(* IEC 61131-3 sources: daoli-st-library/DL_Process (part 39) *)

(* ---- FB_DL_LabelWeekCode.st ---- *)
(*
  Name        : FB_DL_LabelWeekCode
  Category    : DL_Process
  Version     : 1.0.0
  Purpose     : 标签周码/批码打印窗：由年 + 年内日序折算 YYWW 周码，打印请求沿在打印机就绪时发出打印脉冲并锁存周码至请求撤除；/ Label week-code print window: derives a YYWW week code from year and day-of-year, issues a print pulse on request edge when the printer is ready, and latches the code until the request clears
  溯源        : 借 ROADMAP P2（WeekOfYearCalc/DateCoderSync 口径复用），clean-room 实现
  Boundary    : ① 组态闸：年份域 2020..2099 / 年内日序域 1..366 / 打印窗长 > 0 → 锁存故障；
                ② 周码折算：周数 = TRUNC((年内日序 - 1) / 7) + 1（1..53，除子为常量 7，无运行期除零）；
                ③ 打印脉冲 _bPrnC 内部置位 → 段 5 统一出口映射单拍（R187），CASE 内不直写；
                ④ 打印窗计时用 TON 串 ePrint 相位闸（族③），段 0 无 IF 包裹；
                ⑤ nWeekCode 在 eDone 相保持（锁存副本），bPrintReq 撤除沿才回落（族② 保持语义）；
                ⑥ 本件只产生码与脉冲，不驱动打印头（属主边界）。
*)
TYPE E_DL_LwcState :
(
    eIdle  := 0,                             (* 未使能 / Disabled *)
    eReady := 10,                            (* 就绪：等待打印请求（已算码） / Ready *)
    ePrint := 20,                            (* 打印窗进行中 / Printing window *)
    eDone  := 30,                            (* 打印完成（保持周码） / Done, code held *)
    eFault := 90                             (* 故障锁存相 / Fault latched *)
);
END_TYPE

TYPE E_DL_LwcCause :
(
    eNone       := 0,                        (* 无故障成因 / No cause *)
    eCfgIllegal := 1,                        (* 组态非法：年份/日序/窗长越域 / Illegal config *)
    ePhaseBad   := 2                         (* 非法相位兜底 / Illegal phase fallback *)
);
END_TYPE

FUNCTION_BLOCK FB_DL_LabelWeekCode
VAR_INPUT
    nYear     : INT := 2026;                 (* 当前年份，域 2020..2099 [年] / Current year, 2020..2099 *)
    nDayOfYear: INT := 1;                    (* 年内日序（1..366），域 1..366 [日] / Day of year, 1..366 *)
    bPrintReq : BOOL := FALSE;               (* 打印请求电平（上升沿发起）[-] / Print request level *)
    bPrnReady : BOOL := FALSE;               (* 打印机就绪电平 [-] / Printer ready level *)
    tWinLen   : TIME := T#500MS;             (* 打印脉冲窗长，域 > T#0S [ms] / Print pulse window, > 0 *)
    bEnable   : BOOL := TRUE;                (* 使能 [-] / Enable *)
    bReset    : BOOL := FALSE;               (* 复位命令，上升沿清周码与故障 [-] / Reset command *)
END_VAR
VAR_OUTPUT
    nWeekCode : INT;                         (* YYWW 周码（eDone 相保持；低 2 位周数、高位年份后两位）[-] / YYWW week code, held *)
    nWeekNo   : INT;                         (* 年内周数 1..53 [周] / Week number, 1..53 *)
    bPrintPuls: BOOL;                        (* 打印脉冲（窗长电平，tWinLen 定义宽度）[-] / Print pulse level over window *)
    bCodeValid: BOOL;                        (* 周码有效电平（eDone 相为 TRUE）[-] / Code-valid level *)
    eState    : E_DL_LwcState;               (* 状态出口 / State outlet *)
    eCause    : E_DL_LwcCause;               (* 故障成因出口（R190 归因唯一） / Fault cause outlet *)
    bError    : BOOL;                        (* 故障锁存标志 [-] / Fault latch flag *)
END_VAR
VAR
    _eState  : E_DL_LwcState := E_DL_LwcState.eIdle;     (* 内部相位（CASE 唯一写入目标） / Internal phase *)
    _eCause  : E_DL_LwcCause := E_DL_LwcCause.eNone;     (* 故障成因锁存量 / Latched cause *)
    rtReq    : R_TRIG;                       (* 打印请求沿实例，段 0 无条件调用 / Request edge instance *)
    rtReqOff : R_TRIG;                       (* 请求撤除沿实例，段 0 无条件调用 / Request-clear edge instance *)
    rtReset  : R_TRIG;                       (* 复位沿实例，段 0 无条件调用 / Reset edge instance *)
    tonWin   : TON;                          (* 打印脉冲窗计时器（IN 串 ePrint 相位） / Print window timer *)
    _bFault  : BOOL;                         (* 故障锁存位 / Latched fault bit *)
    _bCfgBad : BOOL;                         (* 组态非法当拍量 / Illegal config this scan *)
    _bPrnC   : BOOL;                         (* 打印脉冲窗电平内部量（出口统一映射，R187） / Print-pulse internal level *)
    _nWeekI  : INT;                          (* 周数中间量（折算）[周] / Week number intermediate *)
    _nCodeI  : INT;                          (* 周码中间量（YYWW）[-] / Week code intermediate *)
END_VAR
VAR CONSTANT
    DL_LWC_YMIN  : INT := 2020;              (* 年份域下限 [年] / Year domain floor *)
    DL_LWC_YMAX  : INT := 2099;              (* 年份域上限（YY 码两位十进制安全域）[年] / Year domain ceiling *)
    DL_LWC_DMAX  : INT := 366;               (* 年内日序域上限（含闰年）[日] / Day-of-year domain ceiling *)
    DL_LWC_WMAX  : INT := 53;                (* 周数域上限（折算自洽校验用）[周] / Week number ceiling *)
    DL_LWC_SEVEN : INT := 7;                 (* 周折算除子（常量，无运行期除零）[日/周] / Week divisor *)
    DL_LWC_HUND  : INT := 100;               (* YYWW 折算乘数（常量）[-] / YYWW multiplier *)
END_VAR

(* —— 段 0：当拍判据派生 + 实例无条件刷新（R228A；R_TRIG/TON 全在段 0，无 IF 包裹） —— *)
_bCfgBad := (nYear < DL_LWC_YMIN) OR (nYear > DL_LWC_YMAX)                     (* 年份域闸 / Year gate *)
            OR (nDayOfYear < 1) OR (nDayOfYear > DL_LWC_DMAX)                  (* 日序域闸 / Day-of-year gate *)
            OR NOT (tWinLen > T#0S);                                           (* 窗长正域闸 / Window gate *)
rtReq(CLK := bPrintReq);                                                       (* 请求沿每拍必调 / Request edge every scan *)
rtReqOff(CLK := NOT bPrintReq);                                                (* 请求撤除沿每拍必调 / Request-clear edge every scan *)
rtReset(CLK := bReset);                                                        (* 复位沿每拍必调 / Reset edge every scan *)
tonWin(IN := (_eState = E_DL_LwcState.ePrint) AND bPrintReq, PT := tWinLen);   (* 打印窗计时（串 ePrint 相位闸，族③） / Print timer with phase gate *)

(* —— 段 1：单拍量预清零（R107） —— *)
_bPrnC := FALSE;                                                               (* 打印脉冲内部量预清 / Print-pulse preset *)
bPrintPuls := FALSE;                                                           (* 打印脉冲出口预清 / Print-pulse outlet preset *)
bCodeValid := FALSE;                                                           (* 码有效电平预清 / Code-valid preset *)
_nWeekI := 0;                                                                  (* 周数中间量预清 / Week intermediate preset *)
_nCodeI := 0;                                                                  (* 码中间量预清 / Code intermediate preset *)

(* —— 段 2：复位沿处理（作用域：清故障 + 清周码 + 迁 eIdle，R283 逐项声明） —— *)
IF rtReset.Q THEN
    _bFault := FALSE;                                                          (* 清故障锁存 / Clear fault *)
    _eCause := E_DL_LwcCause.eNone;                                            (* 清成因 / Clear cause *)
    nWeekCode := 0;                                                            (* 清周码出口 / Clear code outlet *)
    nWeekNo := 0;                                                              (* 清周数出口 / Clear week outlet *)
    bCodeValid := FALSE;                                                       (* 清码有效电平 / Clear validity level *)
    _eState := E_DL_LwcState.eIdle;                                            (* 迁未使能相 / Back to idle *)
END_IF

(* —— 段 3：组态故障锁存（锁存至复位沿，R189） —— *)
IF _bCfgBad AND NOT _bFault THEN
    _bFault := TRUE;                                                           (* 锁存故障位 / Latch fault *)
    _eCause := E_DL_LwcCause.eCfgIllegal;                                      (* 成因：组态非法 / Cause: illegal config *)
    _eState := E_DL_LwcState.eFault;                                           (* 同步迁故障相 / Migrate to fault *)
END_IF

(* —— 段 4：CASE 主状态机（ELSE 兜底迁 eFault，红线 6） —— *)
CASE _eState OF
    E_DL_LwcState.eIdle:                                                       (* 未使能：出口确定值 / Disabled *)
        nWeekCode := 0;                                                        (* 失能清周码出口 / Clear code outlet *)
        nWeekNo := 0;                                                          (* 失能清周数出口 / Clear week outlet *)
        bCodeValid := FALSE;                                                   (* 失能清码有效电平 / Clear validity level *)
        IF bEnable AND NOT _bFault THEN
            _eState := E_DL_LwcState.eReady;                                   (* 使能进入就绪 / Enter ready *)
        END_IF
    E_DL_LwcState.eReady:                                                      (* 就绪相：折算周码待打印请求 / Ready *)
        IF NOT bEnable THEN
            _eState := E_DL_LwcState.eIdle;                                    (* 失能回未使能 / Back to idle *)
        ELSE
            _nWeekI := TRUNC(INT_TO_REAL(nDayOfYear - 1) / INT_TO_REAL(DL_LWC_SEVEN)) + 1;   (* 周数折算 = TRUNC((日序-1)/7)+1（除子常量，边界②） / Week number derivation *)
            IF _nWeekI > DL_LWC_WMAX THEN
                _nWeekI := DL_LWC_WMAX;                                        (* 周数上限饱和（最后一次写） / Week ceiling, last write *)
            END_IF
            nWeekNo := _nWeekI;                                                (* 周数出口 / Week outlet *)
            _nCodeI := (nYear MOD DL_LWC_HUND) * DL_LWC_HUND + _nWeekI;        (* YYWW 码 = (年 MOD 100)×100 + 周（乘除均为常量） / YYWW code *)
            nWeekCode := _nCodeI;                                              (* 周码出口（就绪相即为当前码） / Code outlet *)
            IF rtReq.Q AND bPrnReady THEN                                      (* 请求沿 + 就绪：发起打印 / Request edge with ready *)
                _bPrnC := TRUE;                                                (* 打印脉冲内部置位（出口统一映射，R187） / Print-pulse internal *)
                _eState := E_DL_LwcState.ePrint;                               (* 进打印窗相 / To printing *)
            END_IF
        END_IF
    E_DL_LwcState.ePrint:                                                       (* 打印窗相：脉冲电平保持窗长 / Printing *)
        IF NOT bEnable THEN
            _eState := E_DL_LwcState.eIdle;                                    (* 失能回未使能 / Back to idle *)
        ELSE
            _bPrnC := TRUE;                                                    (* 打印窗内脉冲电平保持（窗长由 tonWin 定义） / Pulse level held over window *)
            bCodeValid := TRUE;                                                (* 打印期码有效电平 / Validity level during print *)
            IF rtReqOff.Q THEN                                                 (* 请求撤除沿：提前结束窗 / Request cleared: end window *)
                _eState := E_DL_LwcState.eDone;                                (* 迁完成相（保持周码） / To done *)
            ELSIF tonWin.Q THEN                                                (* 窗长到点：打印完成 / Window elapsed: done *)
                _eState := E_DL_LwcState.eDone;                                (* 迁完成相 / To done *)
            END_IF
        END_IF
    E_DL_LwcState.eDone:                                                       (* 完成相：保持周码至请求撤除后的新请求（族② 保持语义） / Done: hold code *)
        IF NOT bEnable THEN
            _eState := E_DL_LwcState.eIdle;                                    (* 失能回未使能 / Back to idle *)
        ELSIF rtReq.Q THEN                                                     (* 新打印请求沿：重新折算再打印 / New request: re-derive and print *)
            _eState := E_DL_LwcState.eReady;                                   (* 回就绪相重折算 / Back to ready *)
        END_IF
    E_DL_LwcState.eFault:                                                      (* 故障相：冻结保持末值，仅复位沿出 / Fault *)
        ;                                                                      (* 锁存回放（R28） / Replay from latch *)
    ELSE                                                                       (* 非法相位兜底迁安全态 / Illegal phase fallback *)
        _eState := E_DL_LwcState.eFault;                                       (* 迁故障相 / To fault *)
        _bFault := TRUE;                                                       (* 同步锁存 / Latch *)
        _eCause := E_DL_LwcCause.ePhaseBad;                                    (* 成因：非法相位 / Cause: illegal phase *)
END_CASE

(* —— 段 5：出口映射（内部 _b* → 输出，R187；名实双出口，R191） —— *)
bPrintPuls := _bPrnC;                                                          (* 打印脉冲单拍出口 / Print-pulse single-scan outlet *)
bCodeValid := bCodeValid OR (_eState = E_DL_LwcState.eDone);                   (* 码有效电平（打印期与保持期均为 TRUE，族②） / Validity level held in done *)
bError := _bFault;                                                             (* 故障标志镜像 / Fault flag mirror *)
eState := _eState;                                                             (* 状态出口 / State outlet *)
eCause := _eCause;                                                             (* 成因出口 / Cause outlet *)
END_FUNCTION_BLOCK

(* ---- FB_DL_LamEvaGelContent.st ---- *)
(*==============================================================================
 * 组件名称 (Component)  : FB_DL_LamEvaGelContent
 * 所属子库 (Sublibrary) : DL_Process
 * 当前版本 (Version)    : 1.0.0
 * 兼容性 (Platform)     : CODESYS 3.5+ / TwinCAT 3 / 汇川 InoProShop / 施耐德 Machine Expert
 *                         仅依赖 Standard.library（R_TRIG / ABS），零厂商私有库
 * 功能描述 (Function)   : 层压 EVA 交联度估算与合格窗判定。三段工艺换算：
 *                         ① 温度-时间积分 ∫max(0, T - Tref)dt（有效热剂量，
 *                         [°C·min]）；② 线性标定曲线 gel = fGelBase + fKRate·
 *                         Dose（[%]）；③ 合格窗 [fGelLo, fGelHi] 判定。层压
 *                         运行电平控制积分启停。与 Integrator（纯积分）分工：
 *                         本件是积分→标定→判窗三段工艺换算。
 * 来源标签 (Origin)     : ROADMAP §19.2 R12 池（L814），自研 clean-room
 * 边界语义 (Boundary)   : ① 首扫初始化 _bInit（R310：积分类件首拍清剂量）；
 *                         ② 温度 NaN/Inf 拍冻结积分（不累计不判窗）；
 *                         ③ 交联度换算后域钳 [0, 100]（标定外推过冲钳位）；
 *                         ④ 组态闸：基准温度/速率/窗界/扫描秒值域检查 → 故障。
 * 输出语义 (Fallback)   : 【R191】bEnable = FALSE → 积分冻结保持（剂量与交联
 *                         度为资产属性）；eFault 相 → 冻结 + bError = TRUE。
 * 码位     (Codes)      : 按 R297 范式零 16# 码位硬编码；错误出口 BOOL+ENUM(eCause)。
 * 红线自检 (Redline)    : 7 项红线已自检：R1 零全局 ✓｜R2 零物理地址 ✓｜R3 纯 IEC ✓
 *                         R4 除零无涉/NaN 冻结/钳位/组态闸 ✓｜R5 双语同行注释 ✓
 *                         R6 CASE 带 ELSE 兜底迁 eFault ✓｜R7 R_TRIG 段 0 无条件刷新 ✓
 * 验收向量 (Acceptance) : V1 T=150 恒定、Tref=140、fScanS=1.0、fKRate=0.02：
 *                         600 s 后 Dose = 600·10/60 = 100 [°C·min]，
 *                         gel = 基准 20 + 0.02·100 = 22.0 [%]；
 *                         V2 T <= Tref 全程 → Dose=0，gel=基准（不超下界）；
 *                         V3 gel > 100 外推过冲 → 钳 100（边界③）。
 * 修订历史 (Revision)   : 2026-11-20  v1.0.0  R51 首版（批 2 · 序号 10）
 *==============================================================================*)
TYPE E_DL_LgcState :
(
    eIdle  := 0,                             (* 待使能 / Idle *)
    eCalc  := 10,                            (* 积分与判窗运行 / Calc run *)
    eFault := 90                             (* 故障锁存相 / Fault latched phase *)
);
END_TYPE

TYPE E_DL_LgcCause :
(
    eNone       := 0,                        (* 无故障成因 / No cause *)
    eCfgIllegal := 1,                        (* 组态非法：基准/速率/窗界越域 / Illegal config *)
    ePhaseBad   := 2                         (* 非法相位兜底 / Illegal phase fallback *)
);
END_TYPE

FUNCTION_BLOCK FB_DL_LamEvaGelContent
VAR_INPUT
    fTempC    : LREAL := 25.0;               (* 层压温度 [°C] / Lamination temperature *)
    fTempRef  : LREAL := 140.0;              (* 交联基准温度（低于不累计），域 > 0 [°C] / Reference temperature *)
    fKRate    : LREAL := 0.02;               (* 标定斜率，域 > 0 [%/(°C·min)] / Calibration rate *)
    fGelBase  : LREAL := 20.0;               (* 交联度基准截距，域 [0,100] [%] / Base gel content *)
    fGelLo    : LREAL := 75.0;               (* 合格窗下限，域 < fGelHi [%] / Gel window lower *)
    fGelHi    : LREAL := 95.0;               (* 合格窗上限，域 > fGelLo [%] / Gel window upper *)
    fScanS    : LREAL := 1.0;                (* 扫描周期秒值，域 > 1E-6 [s] / Scan period seconds *)
    bProcRun  : BOOL := FALSE;               (* 层压运行电平（积分启停）[-] / Process run level *)
    bEnable   : BOOL := TRUE;                (* 使能 [-] / Enable *)
    bReset    : BOOL := FALSE;               (* 复位命令，上升沿清剂量与输出 [-] / Reset command *)
END_VAR
VAR_OUTPUT
    fDose     : LREAL;                       (* 有效热剂量 [°C·min] / Effective thermal dose *)
    fGelPct   : LREAL;                       (* 交联度估算（钳 0..100）[%] / Gel content estimate *)
    bGelOk    : BOOL;                        (* 合格窗判定（窗口内）[-] / Gel-in-window verdict *)
    eState    : E_DL_LgcState;               (* 状态出口 / State outlet *)
    eCause    : E_DL_LgcCause;               (* 故障成因出口 / Fault cause outlet *)
    bError    : BOOL;                        (* 故障锁存标志 [-] / Fault latch flag *)
END_VAR
VAR
    _eState  : E_DL_LgcState := E_DL_LgcState.eIdle;      (* 内部相位（CASE 唯一写入目标） / Internal phase *)
    _eCause  : E_DL_LgcCause := E_DL_LgcCause.eNone;      (* 故障成因锁存量 / Latched cause *)
    rtReset  : R_TRIG;                       (* 复位沿实例，段 0 无条件调用 / Reset edge instance *)
    _fDose   : LREAL;                        (* 剂量积分锁存 [°C·min] / Dose integrator latch *)
    _fGel    : LREAL;                        (* 交联度派生量 [%] / Gel derived *)
    _bTempBad: BOOL;                         (* 温度非有限当拍量 [-] / Non-finite temperature *)
    _bInit   : BOOL := FALSE;                (* 首扫初始化标志（R310）[-] / First-scan init flag *)
    _bFault  : BOOL;                         (* 故障锁存位 / Latched fault bit *)
    _bCfgBad : BOOL;                         (* 组态非法当拍量 / Illegal config this scan *)
END_VAR
VAR CONSTANT
    DL_LGC_EPS : LREAL := 1.0E-6;            (* 秒值判零容差 [s] / Seconds epsilon *)
    DL_LGC_MIN : LREAL := 60.0;              (* 秒 → 分换算常量 [s/min] / Seconds per minute *)
    DL_LGC_GMAX: LREAL := 100.0;             (* 交联度物理上限 [%] / Gel physical max *)
    DL_LGC_INF : LREAL := 1.0E30;            (* Inf 差判兜底量纲界 [—] / Inf diff guard *)
END_VAR

(* —— 段 0：当拍判据派生 + 实例无条件刷新（R228A） —— *)
_bCfgBad := (fTempRef <= 0.0) OR (fKRate <= 0.0) OR (fGelBase < 0.0) OR (fGelBase > DL_LGC_GMAX)
            OR (fGelLo >= fGelHi) OR (fScanS <= DL_LGC_EPS);   (* 组态闸（R151 全引脚 + 窗界序） / Config gate *)
rtReset(CLK := bReset);                      (* 复位沿每拍必调 / Reset edge every scan *)
_bTempBad := (fTempC <> fTempC) OR ((fTempC - fTempC) <> (fTempC - fTempC))
            OR (ABS(fTempC) > DL_LGC_INF);   (* 温度 NaN 自反 + Inf 差判 + 量纲兜底 / Non-finite temperature *)

(* —— 段 1：首扫初始化（R310：积分类件首拍清剂量，与复位沿同款） —— *)
IF NOT _bInit THEN
    _fDose := 0.0;                           (* 首拍剂量清零 / First-scan dose clear *)
    _fGel := fGelBase;                       (* 首拍交联度取基准 / First-scan gel base *)
    _bInit := TRUE;                          (* 置初始化完成 / Set init done *)
END_IF
_fGel := 0.0;                                (* 交联度当拍量预清（每拍全路径派生，R285） / Gel preset *)
bGelOk := FALSE;                             (* 判窗预清（全路径赋值） / Verdict preset *)

(* —— 段 2：复位沿处理（作用域：清故障 + 清剂量积分 + 清输出 + 迁 eIdle，R283 逐项声明） —— *)
IF rtReset.Q THEN
    _bFault := FALSE;                        (* 清故障锁存 / Clear fault *)
    _eCause := E_DL_LgcCause.eNone;          (* 清成因 / Clear cause *)
    _fDose := 0.0;                           (* 清剂量积分 / Clear dose *)
    fDose := 0.0;                            (* 清剂量出口 / Clear dose outlet *)
    fGelPct := fGelBase;                     (* 交联度回基准 / Gel back to base *)
    _eState := E_DL_LgcState.eIdle;          (* 迁待机相 / Back to idle *)
END_IF

(* —— 段 3：组态闸故障锁存（R45 配对；锁存至复位沿，R189） —— *)
IF _bCfgBad AND NOT _bFault THEN
    _bFault := TRUE;                         (* 锁存故障位 / Latch fault *)
    _eCause := E_DL_LgcCause.eCfgIllegal;    (* 成因：组态非法 / Cause: illegal config *)
    _eState := E_DL_LgcState.eFault;         (* 同步迁故障相 / Migrate to fault *)
END_IF

(* —— 段 4：CASE 主状态机（ELSE 兜底迁 eFault，红线 6） —— *)
CASE _eState OF
    E_DL_LgcState.eIdle:                     (* 待机相 / Idle *)
        IF bEnable AND NOT _bFault AND NOT _bTempBad THEN
            _eState := E_DL_LgcState.eCalc;  (* 进入计算 / Enter calc *)
        END_IF
    E_DL_LgcState.eCalc:                     (* 计算相：积分 + 标定 + 判窗 / Calc *)
        IF NOT bEnable THEN
            _eState := E_DL_LgcState.eIdle;  (* 失能回待机（剂量冻结保持，R191 声明） / Back to idle, dose held *)
        ELSIF bProcRun AND (NOT _bTempBad) THEN   (* 运行电平 + 温度有限才积分 / Integrate when running *)
            IF fTempC > fTempRef THEN        (* 有效热剂量：仅高于基准累计 / Dose above reference *)
                _fDose := _fDose + (fTempC - fTempRef) * fScanS / DL_LGC_MIN;   (* 增量 = ΔT·dt/60 [°C·min]，除子常量 60 无除零 / Dose increment *)
            END_IF
        END_IF                               (* 温度坏值/停运拍：积分冻结（边界②） / Freeze on bad temp *)
        _fGel := fGelBase + fKRate * _fDose; (* 标定曲线换算（乘法无除零） / Calibration transform *)
        IF _fGel < 0.0 THEN
            _fGel := 0.0;                    (* 下界钳位 / Lower clamp *)
        ELSIF _fGel > DL_LGC_GMAX THEN
            _fGel := DL_LGC_GMAX;            (* 上界钳位（外推过冲兜底，边界③） / Upper clamp *)
        END_IF
        IF (_eState = E_DL_LgcState.eCalc) AND (NOT _bTempBad) THEN   (* 判窗仅运行域有效拍 / Verdict in valid scans *)
            fDose := _fDose;                 (* 剂量出口刷新 / Dose outlet *)
            fGelPct := _fGel;                (* 交联度出口刷新 / Gel outlet *)
            IF _fGel < fGelLo THEN
                bGelOk := FALSE;             (* 低于窗 / Below window *)
            ELSIF _fGel > fGelHi THEN
                bGelOk := FALSE;             (* 高于窗 / Above window *)
            ELSE
                bGelOk := TRUE;              (* 窗内（IF 链带 ELSE 兜底，R285） / In window *)
            END_IF
        END_IF
    E_DL_LgcState.eFault:                    (* 故障相：冻结保持，仅复位沿出 / Fault *)
        ;                                    (* 锁存回放（R28） / Replay from latch *)
    ELSE                                     (* 非法相位兜底迁安全态 / Illegal phase fallback *)
        _eState := E_DL_LgcState.eFault;     (* 迁故障相 / To fault *)
        _bFault := TRUE;                     (* 同步锁存 / Latch *)
        _eCause := E_DL_LgcCause.ePhaseBad;  (* 成因：非法相位 / Cause: illegal phase *)
END_CASE

(* —— 段 5：出口映射（bError/eState 同源，R191） —— *)
bError := _bFault;                           (* 故障标志镜像 / Fault flag mirror *)
eState := _eState;                           (* 状态出口 / State outlet *)
eCause := _eCause;                           (* 成因出口 / Cause outlet *)
END_FUNCTION_BLOCK

(* ---- FB_DL_LamHeaterZoneSync.st ---- *)
//==============================================================================
// 功能块：FB_DL_LamHeaterZoneSync ｜ 中文名称：层压机加热板多温区同步跟随
// 所属子库：DL_Process ｜ 版本：v1.0.0 ｜ 兼容：CODESYS V3.5+ / TwinCAT 3 / 汇川 InoProShop
// 功能描述：层压机加热板多温区同步监视——计算有效温区两两最大区差与
//           最差温差对，区差超阈值经确认窗（防瞬态抖动）判失步故障；
//           链速参与跟随语义（链速为 0 时跟随斜率冻结，不除零）。
// 开源溯源 (Origin)：道莅原创实现（参考光伏组件层压机工程惯例 分类与参数域）
// 单位表：T[°C] / 区差[K] / 链速[mm/s] / 确认窗[ms] / 温区下标[区]
// 错误码表：16#0005_01E6 信息级（非有限温区剔除声明，不置 bError）/
//           16#0005_01E7 信息级（区数上限已钳位 8，不置 bError）/
//           16#0005_031E 故障级（区差超限经确认窗确认，置 bError）/
//           16#0005_031F 故障级（有效区数 < 2 无法判区差，置 bError）/
//           16#0005_0320 故障级兜底（置 bError）
// 状态机：N/A（阈值确认窗 + 电平逻辑，无相位状态机；故障经确认窗后以
//           bSyncOk 电平与 031E 表达，原因消失自动恢复，无锁存）
// 边界行为：① 区差 > 阈值持续确认窗 → 故障 031E + bSyncOk := FALSE
//           （R13 AhuDamperStuckDiag 确认窗范式复用）；② 任一温区非有限
//           → 该区剔除出区差统计 + 信息 01E6；有效区数 < 2 → 故障 031F；
//           ③ 链速为 0 → 跟随斜率冻结（不除零），区差统计不受影响；
//           ④ 区数上限钳 8 + 信息 01E7（接口字面量上界 8 与 DL_ZONE_MAX
//           同源，一致性由本件承担验证责任）；⑤ 非使能时输出冻结为零
//           值并 bValid := FALSE（不静默沿用旧差值）。
// 依赖纪律：仅 Standard.library；零跨层调用（两两区差为 O(n²) 遍历的
//           监视语义，非统计算法复制，头注释声明此设计取舍）。
// 修订历史：v1.0.0 2026-11-17 首版（R23 派单 · ROADMAP 光伏 P1 §416）
//==============================================================================

FUNCTION_BLOCK FB_DL_LamHeaterZoneSync
VAR_INPUT
    aZoneTempC    : ARRAY[1..8] OF LREAL;   // 各温区实测 [摄氏度]，下标 1..8，超编路填 0 且不计 / Measured zone temperatures [degC], index 1..8
    uZoneCount    : UINT;                   // 实际温区数 [区]，有效域 0..8，> 8 钳位 / Actual zone count [zones], 0..8, clamped above
    fZoneDiffMaxK : LREAL := 5.0;           // 区差阈值 [K]，须 > 0 / Zone-difference threshold [K], must be > 0
    fBeltSpeedMmS : LREAL;                  // 链速 [毫米/秒]，0 = 停链（跟随冻结） / Belt speed [mm/s], zero = stopped, follow frozen
    bEnable       : BOOL;                   // 使能 [—] / Enable
    bReset        : BOOL;                   // 故障复位 [—]，清除确认窗 / Fault reset, clears the confirm window
END_VAR
VAR_OUTPUT
    fMaxZoneDiffK : LREAL;                  // 当拍最大区差 [K] / Maximum zone difference this scan [K]
    bSyncOk       : BOOL;                   // 同步正常 [—] / Synchronization OK
    uWorstPairA   : UINT;                   // 最大温差对 A 区下标 [区] / Worst pair index A [zone]
    uWorstPairB   : UINT;                   // 最大温差对 B 区下标 [区] / Worst pair index B [zone]
    eErr          : UDINT;                  // 错误码，0 = 无错 / Error code, 0 = no error
    bError        : BOOL;                   // 故障级标志，仅故障级错误置位 / Fault-class flag, set only on fault-level codes
    bValid        : BOOL;                   // 输出可用标志 / Outputs usable flag
END_VAR
VAR
    fbConfirm     : TON;                    // 区差超限确认窗，段 6 无条件刷新 [ms] / Zone-diff confirm window
    _uCountEff    : UINT;                   // 钳位后的生效区数 [区] / Effective clamped zone count
    _uValidZones  : UINT;                   // 非有限剔除后的有效区数 [区] / Valid zone count after culling
    _uI           : UINT;                   // 外层遍历下标 [区] / Outer loop index
    _uJ           : UINT;                   // 内层遍历下标 [区] / Inner loop index
    _fDiff        : LREAL;                  // 当前对区差 [K] / Current pair difference [K]
    _bInit        : BOOL := FALSE;          // 首扫标志，初值 FALSE 取非判定 / First-scan flag, tested negated
    _bCullInfo    : BOOL;                   // 非有限剔除信息当拍标志 / Cull info flag of this scan
    _bClampInfo   : BOOL;                   // 区数钳位信息当拍标志 / Clamp info flag of this scan
    _bIllegal     : BOOL;                   // 非法输入标志（阈值非有限/<= 0） / Illegal input flag
END_VAR
VAR CONSTANT
    DL_ZONE_MAX   : UINT  := 8;             // 温区上限 [区]，与接口字面量上界 8 同源，改动须同步 / Zone ceiling [zones], same source as the literal bound 8, change both together
    DL_LAM_INF    : LREAL := 1.7976931348623157E308; // LREAL 幅值上限 / LREAL magnitude ceiling
    DL_LAM_CONFIRM: TIME  := T#10S;         // 区差超限确认窗 [ms]（R13 范式） / Zone-diff confirm window [ms], R13 pattern
END_VAR

(*------------------------------------------------------------------------------
 * 段 1｜每拍预置：输出先算后出，单拍标志预清零
 *      Outputs computed per scan, one-shot flags pre-cleared
 *-----------------------------------------------------------------------------*)
fMaxZoneDiffK := 0.0;                       // 最大区差预置零 / Max difference preset zero
bSyncOk       := FALSE;                     // 同步正常预置 FALSE / Sync OK preset FALSE
uWorstPairA   := 0;                         // 最差对 A 预置零 / Worst A preset zero
uWorstPairB   := 0;                         // 最差对 B 预置零 / Worst B preset zero
eErr          := 16#0000_0000;              // 错误码每拍重算 / Error code recomputed
bError        := FALSE;                     // 故障标志每拍重算 / Fault flag recomputed
bValid        := FALSE;                     // 可用标志每拍重算 / Usable flag recomputed
_bCullInfo    := FALSE;                     // 剔除信息预清零 / Cull info pre-cleared
_bClampInfo   := FALSE;                     // 钳位信息预清零 / Clamp info pre-cleared
_bIllegal     := FALSE;                     // 非法输入预清零 / Illegal input pre-cleared

(*------------------------------------------------------------------------------
 * 段 2｜首扫初始化
 *      First-scan initialisation
 *-----------------------------------------------------------------------------*)
IF NOT _bInit THEN
    _uCountEff := 0;                        // 生效区数从零起步 / Effective count starts at zero
    _bInit     := TRUE;                     // 首扫只做一次 / The first scan runs once
END_IF

(*------------------------------------------------------------------------------
 * 段 3｜组态与输入防御闸（阈值非法 / 区数钳位）
 *      Configuration and input defense gates
 *-----------------------------------------------------------------------------*)
IF (fZoneDiffMaxK <> fZoneDiffMaxK) OR (ABS(fZoneDiffMaxK) > DL_LAM_INF) OR (fZoneDiffMaxK <= 0.0) THEN
    _bIllegal := TRUE;                      // 阈值非法（031F 无法判差的同类防御，R90 精神） / Illegal threshold
END_IF
IF (fBeltSpeedMmS <> fBeltSpeedMmS) OR (ABS(fBeltSpeedMmS) > DL_LAM_INF) THEN
    _bIllegal := TRUE;                      // 链速非有限防御 / Non-finite belt speed
END_IF
IF uZoneCount > DL_ZONE_MAX THEN
    _uCountEff := DL_ZONE_MAX;              // 区数钳位到 8 / Zone count clamped to 8
    _bClampInfo := TRUE;                    // 钳位信息置位 / Clamp info raised
ELSE
    _uCountEff := uZoneCount;               // 合法区数原值生效 / Valid count applied as-is
END_IF

(*------------------------------------------------------------------------------
 * 段 4｜两两区差扫描（非有限区剔除 + 最差对记录）
 *      Pairwise scan with non-finite culling and worst-pair recording
 *-----------------------------------------------------------------------------*)
_uValidZones := 0;                          // 有效区数清零 / Valid count cleared
FOR _uI := 1 TO _uCountEff DO
    IF _uI <= DL_ZONE_MAX THEN              // 二次闸：越界结构性不可能 / Secondary gate, out-of-bounds impossible
        IF (aZoneTempC[_uI] <> aZoneTempC[_uI]) OR (ABS(aZoneTempC[_uI]) > DL_LAM_INF) THEN
            _bCullInfo := TRUE;             // 非有限区剔除声明 / Non-finite zone culled
        ELSE
            _uValidZones := _uValidZones + 1; // 有效区计数递增 / Valid count increment
        END_IF
        FOR _uJ := _uI + 1 TO _uCountEff DO
            IF _uJ <= DL_ZONE_MAX THEN      // 二次闸 / Secondary gate
                IF (aZoneTempC[_uI] <> aZoneTempC[_uI]) OR (ABS(aZoneTempC[_uI]) > DL_LAM_INF)
                   OR (aZoneTempC[_uJ] <> aZoneTempC[_uJ]) OR (ABS(aZoneTempC[_uJ]) > DL_LAM_INF) THEN
                    (* 任一侧非有限：本对剔除，不计入区差 / Either side non-finite, the pair is culled *)
                    _fDiff := 0.0;          // 本对区差按零计（不参与最差对竞争） / Pair difference counted as zero
                ELSE
                    _fDiff := ABS(aZoneTempC[_uI] - aZoneTempC[_uJ]); // 当前对区差 [K] / Current pair difference [K]
                    IF _fDiff > fMaxZoneDiffK THEN
                        fMaxZoneDiffK := _fDiff; // 更新最大区差 / Update the max difference
                        uWorstPairA := _uI;  // 记录最差对 A / Record worst pair A
                        uWorstPairB := _uJ;  // 记录最差对 B / Record worst pair B
                    END_IF
                END_IF
            END_IF
        END_FOR
    END_IF
END_FOR

(*------------------------------------------------------------------------------
 * 段 5｜确认窗无条件刷新（R40：CASE 之外每拍必调）
 *      Confirm window refreshed unconditionally per R40
 *-----------------------------------------------------------------------------*)
fbConfirm(IN := bEnable AND (NOT _bIllegal) AND (_uValidZones >= 2)
              AND (NOT bReset) AND (fMaxZoneDiffK > fZoneDiffMaxK), PT := DL_LAM_CONFIRM); // 区差超限确认窗（bReset 电平拦截断窗复位） / Zone-diff confirm window, bReset breaks the input to reset

(*------------------------------------------------------------------------------
 * 段 6｜出口与码位（链速为 0 时跟随斜率冻结——本件无斜率输出引脚，
 *       跟随联动由调用方按 fBeltSpeedMmS = 0 自行冻结，边界声明）
 *      Outlet and codes, belt-speed freeze declared for the caller
 *-----------------------------------------------------------------------------*)
IF (NOT bEnable) OR _bIllegal THEN
    bValid := FALSE;                        // 未使能或输入非法：输出不可用 / Not enabled or illegal input, outputs unusable
ELSIF _uValidZones < 2 THEN
    eErr   := 16#0005_031F;                 // 故障级：有效区数 < 2 无法判区差 / Fault: fewer than two valid zones
    bError := TRUE;                         // 置故障标志（R45 配对） / Raise the fault flag
    bValid := FALSE;                        // 输出不可用 / Outputs unusable
ELSIF fbConfirm.Q THEN
    eErr   := 16#0005_031E;                 // 故障级：区差超限经确认窗确认 / Fault: zone difference confirmed
    bError := TRUE;                         // 置故障标志 / Raise the fault flag
    bSyncOk := FALSE;                       // 失步声明 / Desynchronization declared
    bValid := TRUE;                         // 判定结果本身可用 / The verdict itself is usable
ELSE
    bSyncOk := TRUE;                        // 同步正常 / Synchronized
    IF _bCullInfo THEN
        eErr := 16#0005_01E6;               // 信息级：非有限温区已剔除 / Info: non-finite zones culled
    END_IF
    IF _bClampInfo THEN
        eErr := 16#0005_01E7;               // 信息级：区数已钳位 8 / Info: zone count clamped to 8
    END_IF
    bValid := TRUE;                         // 输出可用 / Outputs usable
END_IF
END_FUNCTION_BLOCK

(* ---- FB_DL_LaminatorTempProfile.st ---- *)
(*
  FB_DL_LaminatorTempProfile  —  层压机多温区配方曲线跟随 / Laminator multi-zone temperature profile
  分类 Category : DL_Process
  码位 Code     : 16#06_0_8D
  版本 Version  : 1.0.0
  溯源 Source   : LGF Technology 语义借鉴 · clean-room 实现，仅借分类/参数域/命名，未复制源码
  功能 Function : 1) 每温区按「升温 → 保温 → 降温」三段配方跟随（复用 FB_DL_RampSoakProfile 多实例按温区展开）；
                  2) 全部温区过各自终点窗才置 bProfileDone（单区完成不算完成）；
                  3) 任一温区实测温度无效：该区冻结判定保持末次设定，其余区继续。
  边界 Boundary : ① 段表非法（斜率 <= 0 折算斜坡时间 <= 0、保温时长 < 0、温区数越界）出厂报码；
                  ② 实测温度非有限判 NE43 无效：该温区冻结判定并置信息码，禁塞伪值；
                  ③ 段切换沿冻结一拍防设定阶跃（切换拍不更新区设定输出）；
                  ④ 超时未达窗升级为段故障（锁存），不死等；
                  ⑤ 输出三行同向：区段号 → 区设定 → 完成标志。
  依赖 Depends  : FB_DL_RampSoakProfile × DL_LAM_ZMAX（设定源实例，每拍无条件调用）
  职责边界 Note : 与 FB_DL_CvdTempRamp 同用 RampSoakProfile，但本件面向层压机三段真空/加压
                  配方（段数固定 3、有 bHoldActive 保温保持出口），CVD 件面向多段 Ramp/Soak +
                  均匀性判据，二者行业参数集与判据分立，互不替代。

  码表 Error codes（本件子码步进 16#10，避让邻件码位）:
    16#0002_068D 故障级：段表组态非法（温区数越界 / 斜坡或保温时长 < 0 / 目标温度非有限）
    16#0002_069D 故障级：段超时（保温段计时超限时仍未达窗，锁存需复位）
    16#0002_06AD 信息级：某温区实测温度无效，该区判定已冻结（不置 bError）
*)

TYPE E_DL_LtpPhase :
(
    eIdle    := 0,   // 空闲 / Idle
    eRun     := 10,  // 曲线跟随中 / Profile running
    eDone    := 20,  // 全区完成 / All zones done
    eFrozen  := 30,  // 全部温区无效冻结 / All zones frozen by invalid feedback
    eFault   := 90   // 段故障锁定 / Segment fault locked
);
END_TYPE

FUNCTION_BLOCK FB_DL_LaminatorTempProfile
VAR_INPUT
    bStart        : BOOL;                           // 启动指令，上升沿生效 / Profile start, edge
    bHold         : BOOL;                           // 外部保持（暂停整条曲线）/ External hold
    bReset        : BOOL;                           // 复位，上升沿清段故障 / Reset, clears segment fault
    nZoneCount    : INT := 3;                       // 温区数 [区]，1..DL_LAM_ZMAX / Zone count
    aTgtRampC     : ARRAY[1..4] OF REAL;            // 升温段目标 [°C] × 区 / Ramp segment target [degC] per zone
    aTgtSoakC     : ARRAY[1..4] OF REAL;            // 保温段目标 [°C] × 区 / Soak segment target [degC] per zone
    aTgtCoolC     : ARRAY[1..4] OF REAL;            // 降温段目标 [°C] × 区 / Cool segment target [degC] per zone
    aTempActC     : ARRAY[1..4] OF REAL;            // 各温区实测温度 [°C] / Measured zone temperature [degC]
    tRampUp       : TIME := T#600S;                 // 升温段斜坡时间 [s] / Ramp-up duration
    tSoak         : TIME := T#900S;                 // 保温段保持时间 [s] / Soak duration
    tCoolDown     : TIME := T#600S;                 // 降温段斜坡时间 [s] / Cool-down duration
    fEndWinK      : REAL := 3.0;                    // 终点窗半宽 [K]，域 > 0 / End window half width [K]
    fEps          : REAL := 1.0E-6;                 // 浮点判零容差 [1] / Floating zero tolerance
END_VAR
VAR_OUTPUT
    afZoneSpC     : ARRAY[1..4] OF REAL;            // 各温区设定输出 [°C] / Zone setpoint output [degC]
    anZoneSeg     : ARRAY[1..4] OF INT;             // 各温区当前段号 1..3 / Active segment per zone
    bProfileDone  : BOOL;                           // 全部温区过终点窗 / All zones past end window
    bHoldActive   : BOOL;                           // 保温段激活标志（任一区在保温段）/ Any zone in soak segment
    bError        : BOOL;                           // 故障标志，与故障级码配对 / Fault flag paired with fault codes
    uErrorId      : UDINT;                          // 事件码，0 = 无事件 / Event code, 0 = none
    eStateOut     : E_DL_LtpPhase;                  // 状态机当前态，段尾单点映射 / Phase mapped at tail
END_VAR
VAR
    _eState       : E_DL_LtpPhase := E_DL_LtpPhase.eIdle;  // 内部状态 / Internal state
    afbRs         : ARRAY[1..4] OF FB_DL_RampSoakProfile;  // 每温区一条曲线实例（无条件调用）/ Per-zone profile instance
    rtrStart      : R_TRIG;                         // 启动沿 / Start edge
    rtrReset      : R_TRIG;                         // 复位沿 / Reset edge
    abZoneFrozen  : ARRAY[1..4] OF BOOL;            // 温区冻结掩码（实测无效）/ Zone frozen mask
    abZoneDone    : ARRAY[1..4] OF BOOL;            // 温区过终点窗掩码 / Zone end-window mask
    abSegChgPrev  : ARRAY[1..4] OF BOOL;            // 上拍段切换沿（冻结一拍用）/ Previous segment-change edge
    bCfgOk        : BOOL;                           // 组态合法标志 / Configuration valid
    bZoneOk       : BOOL;                           // 本拍温度数组有效（逐区判定）/ Zone validity this scan
    bAnyFrozen    : BOOL;                           // 存在冻结区 / Any zone frozen
    bAllInvalid   : BOOL;                           // 全部温区无效 / All zones invalid
    nZ            : INT;                            // 温区遍历索引 / Zone loop index
    nSegMax       : INT;                            // 全区最大段号（输出口径）/ Max segment across zones
    uFault        : UDINT;                          // 锁存故障码 / Latched fault code
    uInfo         : UDINT;                          // 信息级码 / Information code
    bTonArmed     : BOOL;                           // 段超时定时器装载条件 / Segment timeout arming condition
END_VAR
VAR CONSTANT
    DL_LAM_ZMAX   : INT := 4;                       // 温区数上限 [区] / Zone count upper bound
    DL_LAM_INFMAX : REAL := 1.0E30;                 // 温度有限值幅值上限 [°C] / Temperature finite bound [degC]
END_VAR

(* === 段 0 · 实例刷新 === *)
rtrStart(CLK := bStart);                          // 每拍刷新启动沿
rtrReset(CLK := bReset);                          // 每拍刷新复位沿

(* === 段 1 · 组态闸 === *)
bCfgOk := (nZoneCount >= 1) AND (nZoneCount <= DL_LAM_ZMAX)    // 温区数域闸
          AND (TIME_TO_REAL(tRampUp) > 0.0)                     // 升温时长 > 0（斜率合法性由时长承载）
          AND (TIME_TO_REAL(tCoolDown) > 0.0) AND (TIME_TO_REAL(tSoak) >= 0.0)
          AND (fEndWinK > fEps);                                // 终点窗半宽正域
FOR nZ := 1 TO DL_LAM_ZMAX DO
    bCfgOk := bCfgOk AND (aTgtRampC[nZ] = aTgtRampC[nZ])        // 目标温度 NaN 自反
              AND (aTgtSoakC[nZ] = aTgtSoakC[nZ]) AND (aTgtCoolC[nZ] = aTgtCoolC[nZ])
              AND (ABS(aTgtRampC[nZ]) < DL_LAM_INFMAX)          // 幅值域闸（仅组态域，实测另行判定）
              AND (ABS(aTgtSoakC[nZ]) < DL_LAM_INFMAX) AND (ABS(aTgtCoolC[nZ]) < DL_LAM_INFMAX);
END_FOR
IF NOT bCfgOk THEN
    uFault := 16#0002_068D;                       // 故障级：段表组态非法
END_IF
IF rtrReset.Q AND bCfgOk THEN
    uFault := 16#0000;                            // 复位沿清段故障锁存（解除路径可达）
    FOR nZ := 1 TO DL_LAM_ZMAX DO
        abZoneDone[nZ] := FALSE;                  // 完成掩码同步复位
        abZoneFrozen[nZ] := FALSE;                // 冻结掩码同步复位
    END_FOR
END_IF
uInfo := 16#0000;                                 // 信息码每拍清零

(* === 段 2 · 逐温区实例调用（无条件）与实测域闸 === *)
bAnyFrozen := FALSE;                              // 冻结汇总先清
bAllInvalid := TRUE;                              // 全无效假设先置
FOR nZ := 1 TO DL_LAM_ZMAX DO
    bZoneOk := (aTempActC[nZ] = aTempActC[nZ]) AND (ABS(aTempActC[nZ]) < DL_LAM_INFMAX);  // NaN 自反 + 幅值闸
    IF bZoneOk THEN
        abZoneFrozen[nZ] := FALSE;                // 该区恢复有效
        abZoneDone[nZ] := abZoneDone[nZ] OR (ABS(aTempActC[nZ] - aTgtCoolC[nZ]) <= fEndWinK + fEps);  // 过终点窗判定（保持型）
        afbRs[nZ](bStart := rtrStart.Q,           // 启动沿下发
                  bHold := bHold OR abZoneFrozen[nZ],   // 外部保持或该区无效冻结（实例内冻结计时）
                  fTrackValue := aTempActC[nZ],   // 无效恢复后无扰回投基准
                  bTrack := FALSE,                // 有效区不跟踪（跟踪入口仅供无效恢复衔接）
                  nSegCount := 3,                 // 固定三段：升温/保温/降温
                  aTarget[1] := aTgtRampC[nZ],    // 段 1 目标：升温
                  aTarget[2] := aTgtSoakC[nZ],    // 段 2 目标：保温
                  aTarget[3] := aTgtCoolC[nZ],    // 段 3 目标：降温
                  aRampTime[1] := tRampUp,        // 段 1 斜坡时间
                  aRampTime[2] := T#0S,           // 段 2 阶跃直达保温目标（保温由时长承载）
                  aRampTime[3] := tCoolDown,      // 段 3 斜坡时间
                  aSoakTime[1] := T#0S,           // 升温到位即切段
                  aSoakTime[2] := tSoak,          // 保温时长
                  aSoakTime[3] := T#0S,           // 降温到位即完成
                  bLoopProfile := FALSE,          // 单次配方不循环
                  bReset := rtrReset.Q);          // 复位沿透传
        IF afbRs[nZ].bSegChange THEN
            abSegChgPrev[nZ] := TRUE;             // 段切换沿：下一拍冻结一拍防设定阶跃
        ELSE
            abSegChgPrev[nZ] := FALSE;            // 非切换拍清标记
        END_IF
        IF NOT abSegChgPrev[nZ] THEN
            afZoneSpC[nZ] := afbRs[nZ].fSetpoint; // 非冻结拍：区设定跟随曲线
        END_IF                                    // 冻结拍：保持上拍设定（防阶跃）
        anZoneSeg[nZ] := afbRs[nZ].nSegAct;       // 段号输出
    ELSE
        abZoneFrozen[nZ] := TRUE;                 // 该区判定冻结（不塞伪值）
        uInfo := 16#0002_06AD;                    // 信息级：温区实测无效该区冻结
        afbRs[nZ](bStart := FALSE, bHold := TRUE, bReset := FALSE,   // 实例仍无条件调用：保持态
                  fTrackValue := aTempActC[nZ], bTrack := TRUE,      // 跟踪入口挂无效值会被实例自身域闸拒绝
                  nSegCount := 3, aTarget[1] := aTgtRampC[nZ], aTarget[2] := aTgtSoakC[nZ],
                  aTarget[3] := aTgtCoolC[nZ], aRampTime[1] := tRampUp, aRampTime[2] := T#0S,
                  aRampTime[3] := tCoolDown, aSoakTime[1] := T#0S, aSoakTime[2] := tSoak,
                  aSoakTime[3] := T#0S, bLoopProfile := FALSE);
        anZoneSeg[nZ] := afbRs[nZ].nSegAct;       // 段号照透传（判定冻结但显示不冻结）
    END_IF
    bAnyFrozen := bAnyFrozen OR abZoneFrozen[nZ]; // 汇总冻结
    bAllInvalid := bAllInvalid AND (NOT bZoneOk); // 汇总全无效
END_FOR

(* === 段 3 · 主状态机（ENUM + CASE，含 ELSE 兜底）=== *)
CASE _eState OF
E_DL_LtpPhase.eIdle :
    bProfileDone := FALSE;                        // 空闲未完成
    bHoldActive := FALSE;                         // 空闲无保温
    IF uFault <> 16#0000 THEN
        _eState := E_DL_LtpPhase.eFault;          // 故障优先
    ELSIF bAllInvalid AND bCfgOk THEN
        _eState := E_DL_LtpPhase.eFrozen;         // 全区无效进冻结
    ELSIF (afbRs[1].nSegAct > 0) OR (afbRs[2].nSegAct > 0)
      OR (afbRs[3].nSegAct > 0) OR (afbRs[4].nSegAct > 0) THEN
        _eState := E_DL_LtpPhase.eRun;            // 任一实例段号非零即运行相
    END_IF

E_DL_LtpPhase.eRun :
    nSegMax := 0;                                 // 段号汇总清零
    bHoldActive := FALSE;                         // 保温标志本拍重算
    FOR nZ := 1 TO nZoneCount DO
        IF anZoneSeg[nZ] > nSegMax THEN
            nSegMax := anZoneSeg[nZ];             // 取全区最大段号
        END_IF
        IF anZoneSeg[nZ] = 2 THEN
            bHoldActive := TRUE;                  // 任一区在保温段即置保温标志
        END_IF
        bTonArmed := (anZoneSeg[nZ] = 2) AND (NOT abZoneFrozen[nZ]);   // 保温超时只对有效区计时
        IF bTonArmed AND (afbRs[nZ].fSoakElapsed > TIME_TO_REAL(tSoak) + 10.0) THEN
            uFault := 16#0002_069D;               // 故障级：保温超时仍未达窗（锁存，不死等）
        END_IF
    END_FOR
    IF uFault <> 16#0000 THEN
        _eState := E_DL_LtpPhase.eFault;          // 故障转出
    ELSIF bAllInvalid THEN
        _eState := E_DL_LtpPhase.eFrozen;         // 全区无效转冻结
    ELSE
        bProfileDone := TRUE;                     // 完成假设：逐区复核
        FOR nZ := 1 TO nZoneCount DO
            bProfileDone := bProfileDone AND (abZoneDone[nZ] OR (afbRs[nZ].bDone AND bZoneOk));  // 全区过窗才完成
        END_FOR
        bProfileDone := bProfileDone AND (NOT bAnyFrozen);   // 存在冻结区不出完成
        IF bProfileDone THEN
            _eState := E_DL_LtpPhase.eDone;       // 转完成相
        END_IF
    END_IF

E_DL_LtpPhase.eDone :
    bHoldActive := FALSE;                         // 完成相无保温
    bProfileDone := TRUE;                         // 完成保持（保持型，防同拍抹除）
    IF rtrStart.Q THEN
        bProfileDone := FALSE;                    // 新启动沿重开
        _eState := E_DL_LtpPhase.eRun;            // 回运行相
    END_IF

E_DL_LtpPhase.eFrozen :
    bProfileDone := FALSE;                        // 冻结相不出完成
    IF (NOT bAllInvalid) AND (uFault = 16#0000) THEN
        _eState := E_DL_LtpPhase.eRun;            // 任一区恢复即回运行（解除路径可达）
    END_IF

E_DL_LtpPhase.eFault :
    bHoldActive := FALSE;                         // 故障相无保温
    IF uFault = 16#0000 THEN
        _eState := E_DL_LtpPhase.eIdle;           // 解锁回空闲
    END_IF

ELSE
    _eState := E_DL_LtpPhase.eFault;              // 非法状态拦截
    uFault := 16#0002_068D;                       // 故障级：相 ID 越界复用组态码段
END_CASE

(* === 段 4 · 输出映射 === *)
bError := (uFault <> 16#0000);                    // 故障标志仅由故障级码置位（R45 配对）
IF bError THEN
    uErrorId := uFault;                           // 故障级优先上报
ELSE
    uErrorId := uInfo;                            // 否则上报信息级码
END_IF
eStateOut := _eState;                             // 输出枚举段尾单点映射（N2 规则）
END_FUNCTION_BLOCK

(* ---- FB_DL_LaminatorVacLeakTrend.st ---- *)
(*==============================================================================
 * 组件名称 (Component)  : FB_DL_LaminatorVacLeakTrend
 * 所属子库 (Sublibrary) : DL_Process
 * 当前版本 (Version)    : 1.0.0
 * 兼容性 (Platform)     : CODESYS 3.5 / TwinCAT 3 / 汇川 InoProShop（纯标准元素，零方言）
 * 功能描述 (Function)   : 真空泄漏率趋势诊断。仅在保压段按采样周期求压强上升速率，与
 *                         滑动基线和绝对上限比较：越基线预警、越绝对上限报警。真空**上升**
 *                         （负泄漏）不刷新基线——放气会把基线抬高，真泄漏将永不报警；基线
 *                         未满样本数时绝对报警恒不置位（不给未标定报警）。不做保压段判定
 *                         本身（由引脚注入）、不做抽气曲线包络、不做阀门控制。
 *                         交付门槛：速率换算用时间转换链，须在 CODESYS / TwinCAT / InoProShop
 *                         三平台各编译验证一次。
 * 溯源 (Origin)         : 道莅 clean-room 防御性实现
 * 本文件内含 (Contains) : TYPE E_DL_LeakState / FUNCTION_BLOCK FB_DL_LaminatorVacLeakTrend
 * 依赖 (Depends)        : 无（仅 Standard.library 的 ABS / TIME_TO_LREAL）
 * 红线自检 (Redline)    : 无外部全局变量、无硬件地址直引 ｜ 全变量中英双语同行注释
 *                         采样周期与上限判零防除零 ｜ 速率非有限即跳过并报信息级 ｜ 基线只
 *                         在正泄漏时刷新 ｜ 采样定时器无条件周期刷新 ｜ 枚举显式赋值 ｜ CASE 含 ELSE
 * 错误码表 (Codes)      : 16#0005_0430 就绪（无越限或非保压段）
 *                         16#0005_0431 信息级 基线样本未满，绝对报警暂不置位（不置故障级标志）
 *                         16#0005_0432 故障级 组态非法（上限 ≤0、基线倍率出域、样本数 <3、采样周期出域）
 *                         16#0005_0433 预留：本版不发码（下一轮区间起点，禁止回填）
 *                         16#0005_0434 信息级 速率非有限，本拍跳过（基线不刷新）
 * 修订历史 (Revision)   : 2026-11-17  v1.0.0  首版入库 · R28 · 阶段三批 3
 * 验收向量 (Acceptance) : 正向 1.0→1.05 kPa/60 s（0.05 kPa/min）、上限 0.1 → 不报警
 *                         反向 1.0→1.5 kPa/60 s（0.5 kPa/min）超上限 0.1 → bLeakAlarm；基线
 *                         0.02、当前 0.06（3 倍 > 倍率 1.1）→ bLeakWarn；上限给 0 →
 *                         16#0005_0432；压强给 NaN → 16#0005_0434 且基线不刷新
 *============================================================================*)

(*-----------------------------------------------------------------------------
 * 枚举: E_DL_LeakState（归属本功能块，同文件发布，全库唯一定义）
 *----------------------------------------------------------------------------*)
TYPE E_DL_LeakState :
(
    eWait  := 0,    // 等待：非保压段或首样本未到 / Waiting, not in the hold phase or no first sample yet
    eTrack := 10,   // 跟踪：按采样周期求速率 / Tracking, the rate is computed per sample period
    eFault := 99    // 故障：组态非法锁存 / Fault, the configuration error is latched
);
END_TYPE

FUNCTION_BLOCK FB_DL_LaminatorVacLeakTrend
VAR_INPUT
    bEnable        : BOOL := FALSE;       // 使能 / Enable
    bHoldPhase     : BOOL := FALSE;       // 保压段有效（仅此段计速率） / Hold phase active, the rate is computed here only
    fVac_kPa       : REAL := 1.0;         // 腔体真空 [kPa(abs)] / Chamber vacuum in kilopascal absolute
    tSampleTime    : TIME := T#100MS;     // 采样周期 [ms]，域 10~1000 / Sampling period, domain 10 to 1000 ms
    fLeakRateMax_kPamin : REAL := 0.1;    // 绝对上限 [kPa/min]，域 0.001~10 / Absolute limit, domain 0.001 to 10
    fBaseK         : REAL := 1.5;         // 基线倍率 [—]，域 1.1~5.0 / Baseline multiplier, domain 1.1 to 5.0
    uBaseSamples   : UINT := 5;           // 基线样本数 [个]，域 3~20 / Baseline sample count, domain 3 to 20
END_VAR
VAR_OUTPUT
    fLeakRate_kPamin  : REAL;             // 当前泄漏率 [kPa/min] / Current leak rate
    fLeakBase_kPamin  : REAL;             // 基线泄漏率 [kPa/min] / Baseline leak rate
    bLeakWarn      : BOOL;                // 越基线预警 / Above the baseline
    bLeakAlarm     : BOOL;                // 越绝对上限报警 / Above the absolute limit
    bError         : BOOL;                // 故障级标志，仅故障级码置位 / Fault-class flag, set on fault codes only
    eErr           : UDINT;               // 错误码，段位 16#0005_xxxx / Error code in segment 16#0005_xxxx
END_VAR
VAR
    _eState        : E_DL_LeakState := E_DL_LeakState.eWait; // 当前相位 / Current phase
    _bInit         : BOOL := FALSE;       // 首扫标志，取非判定 / First-scan flag, tested negated
    _bCfgOk        : BOOL;                // 组态合法标志 / Configuration valid flag
    _bHasSample    : BOOL := FALSE;       // 已有上一拍样本标志 / A previous sample exists
    _bFaultLatch   : BOOL := FALSE;       // 组态故障锁存 / Configuration fault latch
    _fPrev_kPa     : REAL := 0.0;         // 上一拍压强 [kPa(abs)] / Previous pressure sample
    _fDelta        : REAL;                // 本拍压强增量 [kPa] / Pressure increment of this scan
    _fMinSpan      : REAL := 0.1;         // 采样周期换算分钟 [min] / Sampling period in minutes
    _afBase        : ARRAY[1..20] OF REAL; // 基线样本环形表 [kPa/min] / Baseline ring buffer
    _uBaseIdx      : UINT := 1;           // 基线下标 / Baseline index
    _uBaseFill     : UINT := 0;           // 基线已填样本数 [个] / Number of baseline samples collected
    _fBaseSum      : REAL := 0.0;         // 基线样本和 [kPa/min] / Baseline sample sum
    _rtrigSample   : R_TRIG;              // 采样节拍上升沿 / Rising edge of the sample tick
    _tonSample     : TON;                 // 采样周期计时（自复位） / Sampling period timer, self resetting
END_VAR
VAR CONSTANT
    DL_LK_READY    : UDINT := 16#0005_0430;  // 就绪码 / Ready code
    DL_LK_BASE_OFF : UDINT := 16#0005_0431;  // 信息级基线未满码 / Info code for an incomplete baseline
    DL_LK_CFG_BAD  : UDINT := 16#0005_0432;  // 故障级组态非法码 / Fault code for bad configuration
    DL_LK_SKIP     : UDINT := 16#0005_0434;  // 信息级速率非有限码 / Info code for a non-finite rate
    DL_LK_SMP_LO   : TIME := T#10MS;         // 采样周期下限 / Sampling period lower bound
    DL_LK_SMP_HI   : TIME := T#1000MS;       // 采样周期上限 / Sampling period upper bound
    DL_LK_RATE_LO  : REAL := 0.001;          // 绝对上限下限 [kPa/min] / Absolute limit lower bound
    DL_LK_RATE_HI  : REAL := 10.0;           // 绝对上限上限 [kPa/min] / Absolute limit upper bound
    DL_LK_BASEK_LO : REAL := 1.1;            // 基线倍率下限 / Baseline multiplier lower bound
    DL_LK_BASEK_HI : REAL := 5.0;            // 基线倍率上限 / Baseline multiplier upper bound
    DL_LK_SMP_MIN  : UINT := 3;              // 基线最少样本数 [个] / Minimum baseline samples
    DL_LK_SMP_MAX  : UINT := 20;             // 基线最多样本数 [个] / Maximum baseline samples
END_VAR

// 段 1｜输出与单拍标志预置
bLeakWarn := FALSE;                                 // 预警标志预清 / Warning flag pre-cleared
bLeakAlarm := FALSE;                                // 报警标志预清 / Alarm flag pre-cleared
bError := FALSE;                                    // 故障标志预清 / Fault flag pre-cleared
eErr := 0;                                          // 错误码预清 / Error code pre-cleared

// 段 2｜采样定时器与沿实例无条件周期刷新（自复位）
_tonSample(IN := bEnable AND bHoldPhase AND (NOT _tonSample.Q), PT := tSampleTime);
_rtrigSample(CLK := _tonSample.Q);                  // 采样节拍沿 / Sample tick edge

// 段 3｜首扫初始化（判据取非，R19）
IF NOT _bInit THEN
    _eState := E_DL_LeakState.eWait;                // 相位待机起步 / Phase starts waiting
    _bInit := TRUE;                                 // 首扫只做一次 / The first scan runs once
END_IF

// 段 4｜组态闸（上限与采样周期判零防除零）
_bCfgOk := NOT ((fLeakRateMax_kPamin <> fLeakRateMax_kPamin) OR ((fLeakRateMax_kPamin - fLeakRateMax_kPamin) <> (fLeakRateMax_kPamin - fLeakRateMax_kPamin)))
        AND (fLeakRateMax_kPamin >= DL_LK_RATE_LO) AND (fLeakRateMax_kPamin <= DL_LK_RATE_HI)
        AND (fBaseK >= DL_LK_BASEK_LO) AND (fBaseK <= DL_LK_BASEK_HI)
        AND (uBaseSamples >= DL_LK_SMP_MIN) AND (uBaseSamples <= DL_LK_SMP_MAX)
        AND (tSampleTime >= DL_LK_SMP_LO) AND (tSampleTime <= DL_LK_SMP_HI);
IF NOT _bCfgOk THEN
    _bFaultLatch := TRUE;                           // 组态故障锁存 / Configuration fault latched
    eErr := DL_LK_CFG_BAD;                          // 故障级：组态非法 / Fault, bad configuration
    bError := TRUE;
    _eState := E_DL_LeakState.eFault;
END_IF
_fMinSpan := TIME_TO_LREAL(tSampleTime) / 60000.0;  // 采样周期换算分钟 [min] / Sampling period in minutes
IF _fMinSpan < 0.00001 THEN
    _fMinSpan := 0.00001;                           // 换算兜底下限 [min] / Conversion lower bound guard
END_IF

// 段 5｜基线未满闸（不给未标定报警）
IF _uBaseFill < uBaseSamples THEN
    eErr := DL_LK_BASE_OFF;                         // 信息级：基线未满，绝对报警暂不置位 / Info, the baseline is incomplete
END_IF

// 段 6｜速率求取（仅保压段 + 采样沿；非有限即跳过，基线不刷新）
CASE _eState OF
    E_DL_LeakState.eWait:
        IF bHoldPhase AND bEnable THEN
            _bHasSample := FALSE;                   // 新保压段：丢弃上一段样本 / New hold phase, drop the previous sample
            _eState := E_DL_LeakState.eTrack;
        END_IF
    E_DL_LeakState.eTrack:
        IF (NOT bHoldPhase) OR (NOT bEnable) THEN
            _bHasSample := FALSE;                   // 保压结束：样本作废 / Hold finished, the sample is dropped
            _eState := E_DL_LeakState.eWait;
        ELSIF _rtrigSample.Q THEN
            IF (fVac_kPa <> fVac_kPa) OR ((fVac_kPa - fVac_kPa) <> (fVac_kPa - fVac_kPa)) THEN
                eErr := DL_LK_SKIP;                 // 信息级：压强非有限，本拍跳过 / Info, the pressure is not finite
            ELSIF _bHasSample THEN
                _fDelta := fVac_kPa - _fPrev_kPa;           // 压强增量（正 = 泄漏上升）[kPa] / Pressure increment, positive means a leak
                fLeakRate_kPamin := (_fDelta / _fMinSpan);  // 泄漏率 [kPa/min] / Leak rate
                IF _fDelta > 0.0 THEN
                    // 正泄漏才刷新基线：真空上升（负泄漏）不刷基线，否则真泄漏永不报警
                    _fBaseSum := _fBaseSum - _afBase[_uBaseIdx];          // 换出最旧样本 [kPa/min] / Remove the oldest sample
                    _afBase[_uBaseIdx] := fLeakRate_kPamin;               // 写入新样本 [kPa/min] / Insert the new sample
                    _fBaseSum := _fBaseSum + fLeakRate_kPamin;            // 样本和更新 [kPa/min] / Update the sum
                    _uBaseIdx := _uBaseIdx + 1;
                    IF _uBaseIdx > DL_LK_SMP_MAX THEN
                        _uBaseIdx := 1;                                   // 环形回卷 / Ring wrap
                    END_IF
                    IF _uBaseFill < uBaseSamples THEN
                        _uBaseFill := _uBaseFill + 1;                     // 已填样本数 +1 [个] / Sample count incremented
                    END_IF
                    IF _uBaseFill > 0 THEN
                        fLeakBase_kPamin := _fBaseSum / UINT_TO_REAL(_uBaseFill);   // 基线均值 [kPa/min] / Baseline mean
                    END_IF
                END_IF
            END_IF
            _fPrev_kPa := fVac_kPa;                 // 样本快照（唯一写点） / Sample snapshot, the single write point
            _bHasSample := TRUE;
        END_IF
    E_DL_LeakState.eFault:
        eErr := DL_LK_CFG_BAD;                      // 故障级：组态非法保持 / Fault, the configuration error is held
        bError := TRUE;
        IF bEnable AND _bCfgOk AND (NOT bHoldPhase) THEN
            _bFaultLatch := FALSE;                  // 组态修正且退出保压后解除 / Released after the configuration is fixed and the hold phase ends
            _eState := E_DL_LeakState.eWait;
        END_IF
    ELSE
        // 非法相位兜底（故障级）
        eErr := DL_LK_CFG_BAD;
        bError := TRUE;
        _eState := E_DL_LeakState.eFault;
END_CASE

// 段 7｜判据比较（基线未满时绝对报警恒 FALSE）
IF _uBaseFill >= uBaseSamples THEN
    IF fLeakRate_kPamin > fLeakRateMax_kPamin THEN
        bLeakAlarm := TRUE;                         // 越绝对上限报警 / Above the absolute limit
    END_IF
END_IF
IF (_uBaseFill >= uBaseSamples) AND (fLeakBase_kPamin > 0.0) THEN
    IF fLeakRate_kPamin > (fLeakBase_kPamin * fBaseK) THEN
        bLeakWarn := TRUE;                          // 越基线倍率预警 / Above the baseline multiplier
    END_IF
END_IF
IF (NOT bLeakAlarm) AND (NOT bLeakWarn) AND (eErr = 0) THEN
    eErr := DL_LK_READY;                            // 无越限回就绪码 / Ready code when nothing exceeds
END_IF
END_FUNCTION_BLOCK

(* ---- FB_DL_LamTempUniformity.st ---- *)
(*
  FB_DL_LamTempUniformity  —  层压板面多测点温度均匀性诊断 / Laminator plate multi-point temperature uniformity diagnostics
  分类 Category : DL_Process
  码位 Code     : 16#06_0_87
  版本 Version  : 1.0.0
  溯源 Source   : LGF Measurement 语义借鉴 · clean-room 实现，仅借分类/参数域/命名，未复制源码
  功能 Function : 1) 多测点（1..8）温度极差与样本标准差双判据诊断板面均匀性；
                  2) 任一测点失效（无效/NaN/域外）从统计中剔除并在掩码标出，绝不以 0 degC 充当有效值；
                  3) 有效测点 < 2 时不出极差结论（单点极差恒 0 会误判均匀），只报信息级码。
  边界 Boundary : ① 测点数 < 2 不出极差结论；
                  ② 任一测点失效从统计剔除并在掩码标出（禁 0 degC 充当有效值）；
                  ③ 均匀性门限按工艺窗口给常量（VAR CONSTANT），禁写裸数值；
                  ④ 结论三行同向：均值 → 极差 → 均匀标志。
  依赖 Depends  : FB_DL_SignalStatistics（极差稳定性趋势统计，每拍无条件调用）

  码表 Error codes（本件子码步进 16#10，避让邻件码位）:
    16#0002_0687 故障级：测点配置越界（nPointCount 不在 1..8）
    16#0002_0697 故障级：有效测点数为 0（全部失效，无法出任何结论）
    16#0002_06A7 信息级：有效测点 < 2，不出极差结论（不置 bError）
*)

TYPE E_DL_LtuPhase :
(
    eIdle    := 0,   // 空闲 / Idle
    eCollect := 10,  // 测点采集 / Point sampling
    eJudge   := 20,  // 判据计算 / Criterion evaluation
    eVerdict := 30,  // 结论输出 / Verdict output
    eFault   := 90   // 故障锁定 / Fault locked
);
END_TYPE

FUNCTION_BLOCK FB_DL_LamTempUniformity
VAR_INPUT
    bEnable      : BOOL;                          // 总使能，FALSE 回空闲 / Master enable
    bSample      : BOOL := TRUE;                  // 采样使能，TRUE 每拍更新结论 / Sampling enable
    bReset       : BOOL;                          // 复位，上升沿清故障与趋势窗 / Reset
    nPointCount  : INT := 4;                      // 测点总数 [点]，域 1~8 / Point count, 1..8
    afTempC      : ARRAY[1..8] OF REAL;           // 各测点温度 [degC]，域 −20~400 / Per-point temperature [degC]
    abPointValid : ARRAY[1..8] OF BOOL;           // 各测点通道有效标志 / Per-point channel valid flag
END_VAR
VAR_OUTPUT
    fMeanC       : REAL;                          // 有效测点温度均值 [degC] / Mean over valid points [degC]
    fRangeC      : REAL;                          // 极差（最大 − 最小）[degC] / Peak-to-peak [degC]
    fStdDevC     : REAL;                          // 样本标准差（n−1）[degC] / Sample standard deviation [degC]
    nValidPts    : INT;                           // 有效测点数 [点] / Valid point count
    abValidMask  : ARRAY[1..8] OF BOOL;           // 有效测点掩码 [开关]，索引 = 物理测点号 / Valid point mask
    bUniform     : BOOL;                          // 均匀合格（极差与标准差双判据均过）/ Uniform, both criteria pass
    bWarn        : BOOL;                          // 均匀性告警（保持型）/ Uniformity warning, held
    bError       : BOOL;                          // 故障标志，与故障级码配对 / Fault flag paired with fault codes
    uErrorId     : UDINT;                         // 事件码，0 = 无事件 / Event code, 0 = none
    eStateOut    : E_DL_LtuPhase;                 // 状态机当前态，段尾单点映射 / Phase mapped at tail
END_VAR
VAR
    _eState      : E_DL_LtuPhase := E_DL_LtuPhase.eIdle;  // 内部状态 / Internal state
    rtrReset     : R_TRIG;                        // 复位沿 / Reset edge
    statRange    : FB_DL_SignalStatistics;        // 极差趋势统计（无条件调用）/ Range trend statistics
    nN           : INT;                           // 钳位后测点数 [点] / Clamped point count
    nI           : INT;                           // 测点循环下标 / Point loop index
    nValid       : INT;                           // 有效测点计数 [点] / Valid point counter
    fSum         : REAL;                          // 温度和 [degC] / Temperature sum [degC]
    fMin         : REAL;                          // 有效最小值 [degC] / Valid minimum [degC]
    fMax         : REAL;                          // 有效最大值 [degC] / Valid maximum [degC]
    fMeanBuf     : REAL;                          // 均值暂存 [degC] / Mean buffer [degC]
    fDevSum      : REAL;                          // 偏差平方和 [degC^2] / Squared deviation sum
    fVar         : REAL;                          // 样本方差 [degC^2] / Sample variance
    bStatOk      : BOOL;                          // 统计量可算标志 / Statistics computable
    uFault       : UDINT;                         // 锁存故障码 / Latched fault code
    uInfo        : UDINT;                         // 信息级码 / Information code
END_VAR
VAR CONSTANT
    DL_LTU_PTMAX   : INT := 8;                    // 测点数组上界 [点] / Point array bound
    DL_LTU_RANGEMAX: REAL := 3.0;                 // 工艺允许极差上限 [degC]（工艺窗口常量）/ Process range limit [degC]
    DL_LTU_STDMAX  : REAL := 1.5;                 // 工艺允许标准差上限 [degC]（工艺窗口常量）/ Process std limit [degC]
    DL_LTU_TMIN    : REAL := -20.0;               // 测点物理域下限 [degC] / Point domain low [degC]
    DL_LTU_TMAX    : REAL := 400.0;               // 测点物理域上限 [degC] / Point domain high [degC]
END_VAR

(* === 段 0 · 实例刷新（无条件周期调用）=== *)
rtrReset(CLK := bReset);                          // 每拍刷新复位沿

(* === 段 1 · 组态闸与测点掩码（失效点剔除，禁 0 degC 充数）=== *)
nN := nPointCount;                                // 测点数取用前钳位
IF nN < 1 THEN
    nN := 1;
END_IF
IF nN > DL_LTU_PTMAX THEN
    nN := DL_LTU_PTMAX;
END_IF
IF (nPointCount < 1) OR (nPointCount > DL_LTU_PTMAX) THEN
    uFault := 16#0002_0687;                       // 故障级：测点配置越界
END_IF
IF rtrReset.Q THEN
    uFault := 16#0000;                            // 复位沿清锁存
    bWarn := FALSE;                               // 告警同步复位
END_IF

(* === 段 2 · 主状态机（ENUM + CASE，含 ELSE 兜底）=== *)
CASE _eState OF
E_DL_LtuPhase.eIdle :
    bStatOk := FALSE;                             // 空闲不可算
    uInfo := 16#0000;                             // 信息码清零
    IF uFault = 16#0002_0687 THEN
        _eState := E_DL_LtuPhase.eFault;          // 组态故障优先
    ELSIF bEnable AND bSample THEN
        _eState := E_DL_LtuPhase.eCollect;        // 进入采集相
    END_IF

E_DL_LtuPhase.eCollect :
    nValid := 0;                                  // 有效点计数清零
    fSum := 0.0;                                  // 温度和清零
    fMin := 1.0E30;                               // 最小值初值取极大
    fMax := -1.0E30;                              // 最大值初值取极小
    FOR nI := 1 TO DL_LTU_PTMAX DO
        IF nI <= nN THEN
            abValidMask[nI] := abPointValid[nI]
                               AND (afTempC[nI] = afTempC[nI])                    // NaN 自反判据
                               AND (ABS(afTempC[nI]) < 1.0E30)                    // Inf 上限兜底
                               AND (afTempC[nI] >= DL_LTU_TMIN)
                               AND (afTempC[nI] <= DL_LTU_TMAX);                  // 物理域闸
            IF abValidMask[nI] THEN
                nValid := nValid + 1;                 // 有效点累加
                fSum := fSum + afTempC[nI];           // 温度和累加
                IF afTempC[nI] < fMin THEN
                    fMin := afTempC[nI];              // 更新最小值
                END_IF
                IF afTempC[nI] > fMax THEN
                    fMax := afTempC[nI];              // 更新最大值
                END_IF
            END_IF
        ELSE
            abValidMask[nI] := FALSE;                 // 超出配置的测点掩码置 FALSE
        END_IF
    END_FOR
    nValidPts := nValid;                          // 有效点输出
    IF nValid >= 1 THEN
        fMeanBuf := fSum / INT_TO_REAL(nValid);   // 均值分母已判 > 0
    ELSE
        fMeanBuf := 0.0;                          // 无效点：均值不出结论
    END_IF
    fMeanC := fMeanBuf;                           // 均值输出
    _eState := E_DL_LtuPhase.eJudge;              // 转判据相

E_DL_LtuPhase.eJudge :
    IF nValidPts >= 2 THEN
        fRangeC := fMax - fMin;                   // 极差：点数 >= 2 才有意义
        fDevSum := 0.0;                           // 偏差平方和清零
        FOR nI := 1 TO DL_LTU_PTMAX DO
            IF (nI <= nN) AND abValidMask[nI] THEN
                fDevSum := fDevSum + (afTempC[nI] - fMeanC) * (afTempC[nI] - fMeanC);   // 逐点累加偏差平方
            END_IF
        END_FOR
        fVar := fDevSum / INT_TO_REAL(nValidPts - 1);   // 样本方差，分母 n−1 >= 1
        IF fVar > 0.0 THEN
            fStdDevC := SQRT(fVar);               // 标准差
        ELSE
            fStdDevC := 0.0;                      // 方差非正：标准差 0
        END_IF
        bStatOk := TRUE;                          // 统计量有效
    ELSE
        fRangeC := 0.0;                           // 点数不足：极差不出结论
        fStdDevC := 0.0;                          // 标准差不出结论
        bStatOk := FALSE;                         // 统计量无效
        uInfo := 16#0002_06A7;                    // 信息级：有效测点 < 2
    END_IF
    _eState := E_DL_LtuPhase.eVerdict;            // 转结论相

E_DL_LtuPhase.eVerdict :
    IF bStatOk THEN
        bUniform := (fRangeC <= DL_LTU_RANGE_MAX + 1.0E-6) AND (fStdDevC <= DL_LTU_STDMAX + 1.0E-6);  // 双判据带容差
        IF NOT bUniform THEN
            bWarn := TRUE;                        // 置位型：均匀性告警（段尾不清零）
        ELSE
            bWarn := FALSE;                       // 恢复均匀即解除告警（可到达的解除路径）
        END_IF
    ELSE
        bUniform := FALSE;                        // 无法判定：不给合格结论
    END_IF
    IF (NOT bEnable) OR rtrReset.Q THEN
        _eState := E_DL_LtuPhase.eIdle;           // 失能/复位回空闲
    ELSIF bSample THEN
        _eState := E_DL_LtuPhase.eCollect;        // 连续采样
    END_IF

E_DL_LtuPhase.eFault :
    bUniform := FALSE;                            // 故障态不给合格结论
    bStatOk := FALSE;                             // 统计无效
    IF uFault = 16#0000 THEN
        _eState := E_DL_LtuPhase.eIdle;           // 解锁回空闲
    END_IF

ELSE
    _eState := E_DL_LtuPhase.eFault;              // 非法状态拦截
    uFault := 16#0002_0697;                       // 故障级：相 ID 越界（枚举兜底路径）
END_CASE

(* === 段 3 · 极差趋势统计实例（每拍无条件调用）=== *)
statRange(fIn := fRangeC,                         // 极差序列
          bSample := bStatOk AND bSample,         // 仅结论有效时采样
          nWindow := 32,                          // 窗口 32 点
          bClear := rtrReset.Q);                  // 复位清窗

(* === 段 4 · 输出映射（三行同向：均值 → 极差 → 均匀标志）=== *)
IF nValidPts = 0 THEN
    uFault := 16#0002_0697;                       // 故障级：全部测点失效，无法出结论
END_IF
bError := (uFault <> 16#0000);                    // 故障标志仅由故障级码置位（R45 配对）
IF bError THEN
    uErrorId := uFault;                           // 故障级优先上报
ELSE
    uErrorId := uInfo;                            // 否则上报信息级码
END_IF
eStateOut := _eState;                             // 输出枚举段尾单点映射（N2 规则）
END_FUNCTION_BLOCK

(* ---- FB_DL_LaserDescumStep.st ---- *)
(*
  组件名 Component   : FB_DL_LaserDescumStep
  子库 Sublibrary    : DL_Process
  版本 Version       : 1.0.0
  兼容性 Platform    : CODESYS 3.5 / TwinCAT 3 / 汇川 InoProShop / Machine Expert（仅 Standard.library）
  功能 Function      : 激光去渣（descum）工步（自研行业池：半导体）：
                       1) 工步参数集：功率/扫速/圈数以输入引脚承载，工步沿启动；
                       2) 逐圈执行：每圈时长 tPassDur，圈计数达到 nPassCount 后停发；
                       3) 终点判据双路：反射率 >= fReflectEndPct 持续 tReflConfirm
                       确认（仪器路）或 bVisConfirm 操作员目视沿（人判路），任一
                       达成即提前结束（早退路径，不发参数变更）；
                       4) 工步超时：tStepTo 专用超时 TON（专用超时件命名），超时即
                       故障锁存（禁把配方时长接到段超时）。
  边界 Boundary      : ① 本件只出激光使能与参数就绪标志，不写物理 IO；
                       ② 工步沿启动后参数集冻结快照（工步中改参不生效，禁中途
                       变参重推断）；圈数域 [1, 99]；
                       ③ 故障锁存解除唯一路径 = bReset 上升沿（输入引脚，恒可达）；
                       ④ 无全局变量引用、无外部变量声明、无物理地址寻址。
  依赖 Depends       : Standard.library（R_TRIG / TON）
  溯源 Origin        : 道莅自研 clean-room（自研行业池：半导体去渣工步共性语义，
                       零外部代码行复制）
  码位 Code          : 16#06_0_C1（Process 段 0006，C 子带 C1 格）
  码表 Error codes（本件格 06_0_C1，单轨子道：故障 0x02C1 / 信息 0x01C1 / 0x03C1）:
    16#0006_02C1 故障级：工步故障总码（工步超时 / 组态非法 / 输入非有限），
                 锁存至复位
    16#0006_01C1 信息级：反射率早退沿（仪器判据达成提前结束拍）
    16#0006_03C1 信息级：目视早退沿（操作员确认提前结束拍）
  修订历史 Revision  :
    2026-11-19  v1.0.0  R44 首版（批次 4 · 序号 18）
*)

TYPE E_DL_LdsPhase :
(
    eIdle  := 0,    // 空闲：等工步沿 / Idle, waiting step edge
    eRun   := 10,   // 工步：逐圈执行 + 终点监视 / Running, pass loop and endpoint watch
    eDone  := 20,   // 完成：工步结论驻留 / Done, step verdict held
    eFault := 90    // 故障：工步锁存 / Fault, latched
);
END_TYPE

FUNCTION_BLOCK FB_DL_LaserDescumStep
VAR_INPUT
    bStartCmd    : BOOL;                   // 工步启动（上升沿承载）[-] / Step start edge
    bReset       : BOOL;                   // 上升沿清故障锁存 [-] / Reset edge
    bVisConfirm  : BOOL;                   // 目视确认（上升沿承载）[-] / Visual confirm edge
    fPowerPct    : REAL := 80.0;           // 激光功率 [%]，域 0..100 / Laser power
    fScanSpeedMmS: REAL := 100.0;          // 扫描速度 [mm/s] / Scan speed
    nPassCount   : INT := 3;               // 计划圈数 [圈]，域 1..99 / Planned pass count
    fReflectPct  : REAL;                   // 反射率实测 [%] / Measured reflectivity
    fReflectEndPct: REAL := 60.0;          // 反射率终点阈 [%] / Reflectivity endpoint threshold
    tPassDur     : TIME := T#10S;          // 每圈时长 [毫秒] / Pass duration
    tReflConfirm : TIME := T#2S;           // 反射率确认窗 [毫秒] / Reflectivity confirm window
    tStepTo      : TIME := T#600S;         // 工步超时 [毫秒] / Step timeout
END_VAR
VAR_OUTPUT
    bLaserEnable : BOOL;                   // 激光使能输出 [-] / Laser enable output
    bParamReady  : BOOL;                   // 参数集就绪标志（工步沿冻结快照有效）[-] / Parameter ready flag
    nPassDone    : INT;                    // 已完成圈数 [圈] / Completed pass count
    bEarlyExit   : BOOL;                   // 早退标志（终点判据提前达成）[-] / Early exit flag
    ePhase       : E_DL_LdsPhase;          // 相位出口，段尾单点映射 / Phase outlet
    bError       : BOOL;                   // 故障锁存标志 [-] / Fault latch flag
    uErrId       : UDINT;                  // 事件码，0 = 无事件 / Event code
END_VAR
VAR
    rtReset   : R_TRIG;                    // 复位沿实例，段 0 无条件刷新 / Reset edge
    rtStart   : R_TRIG;                    // 工步沿实例，段 0 无条件刷新 / Start edge
    rtVisConf : R_TRIG;                    // 目视确认沿实例，段 0 无条件刷新 / Visual confirm edge
    tonPassDur: TON;                       // 每圈计时（独立实例） / Pass duration timer
    tonReflConf: TON;                      // 反射率确认窗 / Reflectivity confirm timer
    tonStepTo : TON;                       // 工步超时（专用超时件命名） / Step timeout
    _ePhase   : E_DL_LdsPhase := E_DL_LdsPhase.eIdle;  // 内部相位（CASE 唯一写入目标）/ Internal phase
    _nPassPlan: INT;                       // 冻结计划圈数 [圈] / Frozen planned passes
    _bFault   : BOOL;                      // 故障锁存位（锁存量） / Latched fault bit
    _uFault   : UDINT;                     // 故障码锁存（锁存量） / Latched fault code
    _bCfgBad  : BOOL;                      // 组态非法当拍量 [-] / Config illegal flag
    _bNonFin  : BOOL;                      // 输入非有限当拍量 [-] / Non-finite input flag
END_VAR
VAR CONSTANT
    DL_PASS_MAX : INT  := 99;              // 圈数上限 [圈] / Pass count ceiling
    DL_PASS_MIN : INT  := 1;               // 圈数下限 [圈] / Pass count floor
    DL_ONE      : INT  := 1;               // 单位圈数常量 [圈] / One pass
    DL_ABS_MAX  : REAL := 1.0E30;          // 有限值判定上界 [工程单位] / Finite bound
    DL_ZERO     : REAL := 0.0;             // 零常量 [工程单位] / Zero constant
END_VAR

(* —— 段 0｜沿与定时器每拍无条件刷新（禁置于 IF/CASE 内） —— *)
rtReset  (CLK := bReset);
rtStart  (CLK := bStartCmd);
rtVisConf(CLK := bVisConfirm);
tonPassDur (IN := (_ePhase = E_DL_LdsPhase.eRun) AND (NOT _bFault), PT := tPassDur);
tonReflConf(IN := (_ePhase = E_DL_LdsPhase.eRun) AND (fReflectPct >= fReflectEndPct)
            AND (NOT _bFault), PT := tReflConfirm);
tonStepTo  (IN := (_ePhase = E_DL_LdsPhase.eRun) AND (NOT _bFault), PT := tStepTo);

(* —— 段 1｜瞬时量预清零（锁存量 _bFault/_uFault/_nPassPlan/bEarlyExit 不入清单） —— *)
uErrId   := 16#0000_0000;
_bCfgBad := FALSE;
_bNonFin := FALSE;

(* —— 段 2｜复位沿：故障一次性清干净，相位回空闲，激光使能撤销 —— *)
IF rtReset.Q THEN
    _bFault := FALSE;
    _uFault := 16#0000_0000;
    bLaserEnable := FALSE;
    bParamReady  := FALSE;
    _ePhase := E_DL_LdsPhase.eIdle;
END_IF

(* —— 段 3｜组态闸与非有限判据 —— *)
IF (fPowerPct <= DL_ZERO) OR (fPowerPct > DL_ABS_MAX) OR (fScanSpeedMmS <= DL_ZERO)
   OR (nPassCount < DL_PASS_MIN) OR (nPassCount > DL_PASS_MAX) OR (tPassDur = T#0S)
   OR (tReflConfirm = T#0S) OR (tStepTo = T#0S) OR (fReflectEndPct <= DL_ZERO) THEN
    _bCfgBad := TRUE;
END_IF
IF (fReflectPct <> fReflectPct) OR ((fReflectPct - fReflectPct) <> DL_ZERO) THEN
    _bNonFin := TRUE;
END_IF

(* —— 段 4｜主状态机：四态全覆盖 + ELSE 兜底 —— *)
CASE _ePhase OF

E_DL_LdsPhase.eIdle:
    bLaserEnable := FALSE;
    IF _bFault THEN
        bError := TRUE;                  // 故障锁存回放（R189）
    END_IF
    IF rtStart.Q AND (NOT _bFault) AND (NOT _bCfgBad) AND (NOT _bNonFin) THEN
        _nPassPlan := nPassCount;        // 参数集冻结快照（工步中改参不生效）
        nPassDone  := 0;
        bEarlyExit := FALSE;
        bParamReady := TRUE;
        bLaserEnable := TRUE;
        _ePhase := E_DL_LdsPhase.eRun;
    ELSIF rtStart.Q AND (_bFault OR _bCfgBad OR _bNonFin) THEN
        _bFault := TRUE;                 // 带病启动拒绝
        _uFault := 16#0006_02C1;
        bError  := TRUE;
        _ePhase := E_DL_LdsPhase.eFault;
    END_IF

E_DL_LdsPhase.eRun:
    bLaserEnable := TRUE;
    IF _bNonFin THEN
        _bFault := TRUE;
        _uFault := 16#0006_02C1;
        bError  := TRUE;
        _ePhase := E_DL_LdsPhase.eFault;
    ELSIF rtVisConf.Q THEN
        bEarlyExit := TRUE;              // 人判路早退：终点判据提前达成
        uErrId := 16#0006_03C1;          // 信息级：目视早退沿
        bLaserEnable := FALSE;
        _ePhase := E_DL_LdsPhase.eDone;
    ELSIF tonReflConf.Q THEN
        bEarlyExit := TRUE;              // 仪器路早退：反射率确认达成
        uErrId := 16#0006_01C1;          // 信息级：反射率早退沿
        bLaserEnable := FALSE;
        _ePhase := E_DL_LdsPhase.eDone;
    ELSIF tonPassDur.Q THEN
        nPassDone := nPassDone + DL_ONE; // 一圈完成：圈计数累加
        IF nPassDone >= _nPassPlan THEN
            bLaserEnable := FALSE;       // 圈数达成：停发（正常收口）
            _ePhase := E_DL_LdsPhase.eDone;
        END_IF
    ELSIF tonStepTo.Q THEN
        _bFault := TRUE;                 // 工步超时（配方时长接段计，超时独立承载）
        _uFault := 16#0006_02C1;
        bError  := TRUE;
        bLaserEnable := FALSE;
        _ePhase := E_DL_LdsPhase.eFault;
    END_IF

E_DL_LdsPhase.eDone:
    bLaserEnable := FALSE;
    IF NOT bStartCmd THEN
        _ePhase := E_DL_LdsPhase.eIdle;  // 工步指令撤销：回空闲（结论锁存保留）
    END_IF

E_DL_LdsPhase.eFault:
    bLaserEnable := FALSE;               // 故障相：激光使能安全侧撤销
    bError := TRUE;
    ;                                    // 故障相驻留：只认复位沿（段 2 迁出）

ELSE
    _bFault := TRUE;                     // 兜底：非法相位锁存
    _uFault := 16#0006_02C1;
    bError  := TRUE;
    _ePhase := E_DL_LdsPhase.eFault;
END_CASE

(* —— 段 5｜相位出口单点映射 —— *)
ePhase := _ePhase;
END_FUNCTION_BLOCK

(* ---- FB_DL_LaserWeldPowerSeq.st ---- *)
(*
  FB_DL_LaserWeldPowerSeq  —  激光焊三段功率斜坡配方序列 / Laser weld three-stage power ramp sequencer
  分类 Category : DL_Process
  码位 Code     : 16#06_0_80
  版本 Version  : 1.0.0
  溯源 Source   : LGF SignalGenerators + LBP 语义借鉴 · clean-room 实现，仅借分类/参数域/命名，未复制源码
  功能 Function : 1) 按「预焊-满焊-收弧」三段配方（功率/速度/离焦）推进时序，每段由独立 TON 计时，计时器在 FB 主体无条件刷新；
                  2) 段切换当拍冻结功率/速度/离焦输出一拍，沿用上一拍指令，防阶跃冲击焊头与熔池；
                  3) 配方越界（功率 <= 0 或 > 额定）走组态闸出厂即锁存报码，不做运行时钳位掩盖。
  边界 Boundary : ① 三段功率/速度域反算见下方「类型可表性」段；
                  ② 段切换当拍冻结输出功率一拍（由 nSegNow 与 nSegPrev 比较实现，无标志位清零覆盖风险）；
                  ③ 配方越界走组态闸锁存报码，禁运行时钳位掩盖；
                  ④ 中止/失能三行同向：功率指令 0 → 段号 0 → 出光标志 FALSE。
  依赖 Depends  : None

  类型可表性（极限值 → 类型可表性反算）:
    额定功率上限 6000.0 W，功率分辨率 0.1 W → 6000.0 / 0.1 = 60000 计数，远小于 REAL 尾数可精确表出的
    整数上限 16777216，故 0.1 W 步进在本件量程内可精确表出，无舍入溢出。
    速度上限 500.000 mm/s，分辨率 0.001 mm/s → 500000 计数，同样可表。
    离焦 ±10.000 mm，分辨率 0.001 mm → 20000 计数，可表。
    结论：本件不做饱和换算，只做域闸判据。

  码表 Error codes（本件子码步进 16#10，避让邻件码位）:
    16#0002_0680 故障级：配方越界（功率/速度/时间/离焦域外）→ 组态闸锁存，需 bReset 上升沿清除
    16#0002_0690 故障级：段序号越界或段驻留时间为 0（枚举兜底路径）
    16#0002_06A0 信息级：段切换冻结拍已发生（诊断用，永不置 bError）
*)

TYPE E_DL_LwpsPhase :
(
    eIdle   := 0,    // 空闲待命 / Idle
    ePrep   := 10,   // 预焊段 / Pre-weld stage
    eFull   := 20,   // 满焊段 / Full-weld stage
    eCrater := 30,   // 收弧段 / Crater fill stage
    eDone   := 40,   // 序列完成 / Sequence done
    eFault  := 90    // 故障锁定 / Fault locked
);
END_TYPE

FUNCTION_BLOCK FB_DL_LaserWeldPowerSeq
VAR_INPUT
    bEnable      : BOOL;                          // 总使能，FALSE 回空闲并清功率 / Master enable
    bStart       : BOOL;                          // 启动指令，上升沿有效 / Start command, rising edge
    bAbort       : BOOL;                          // 中止指令，上升沿回空闲 / Abort command, rising edge
    bReset       : BOOL;                          // 复位指令，上升沿清锁存故障 / Reset command, rising edge
    afSegPowerW  : ARRAY[1..3] OF REAL;           // 三段激光功率配方 [W]，域 0 < P <= fRatedPowerW / Per-stage power [W]
    afSegSpeed   : ARRAY[1..3] OF REAL;           // 三段焊接速度配方 [mm/s]，域 > 0 / Per-stage weld speed [mm/s]
    afSegDefocus : ARRAY[1..3] OF REAL;           // 三段离焦量配方 [mm]，正负双向 / Per-stage defocus [mm]
    atSegTime    : ARRAY[1..3] OF TIME;           // 三段驻留时间 [ms]，域 > 0 / Per-stage dwell time [ms]
    fRatedPowerW : REAL := 6000.0;                // 激光器额定功率 [W]，域 > 0 / Rated laser power [W]
    fDefocusMax  : REAL := 10.0;                  // 离焦允许幅值 [mm]，域 > 0 / Defocus magnitude limit [mm]
    fEps         : REAL := 1.0E-6;                // 浮点判零容差 [1] / Floating zero tolerance
END_VAR
VAR_OUTPUT
    fPowerCmdW   : REAL;                          // 功率指令 [W]，段切换当拍冻结 / Power command [W], frozen on switch
    fSpeedCmd    : REAL;                          // 焊接速度指令 [mm/s] / Weld speed command [mm/s]
    fDefocusCmd  : REAL;                          // 离焦指令 [mm] / Defocus command [mm]
    nSegNow      : INT;                           // 当前段号 1..3，0 = 未运行 / Current stage 1..3, 0 = inactive
    bWeldActive  : BOOL;                          // 出光中标志 / Emission active flag
    bSeqDone     : BOOL;                          // 全序列完成，保持型 / Sequence done, level held
    nFreezeCount : INT;                           // 段切换冻结拍累计 [拍]，钳 32000 / Accumulated freeze scans
    bError       : BOOL;                          // 故障标志，与故障级码配对 / Fault flag paired with fault codes
    uErrorId     : UDINT;                         // 事件码，0 = 无事件 / Event code, 0 = none
    eStateOut    : E_DL_LwpsPhase;                // 状态机当前态，段尾单点映射 / Phase mapped at tail
END_VAR
VAR
    _eState      : E_DL_LwpsPhase := E_DL_LwpsPhase.eIdle; // 内部状态（唯一真值）/ Internal state, single source of truth
    rtrStart     : R_TRIG;                        // 启动沿检测实例 / Start edge instance
    rtrAbort     : R_TRIG;                        // 中止沿检测实例 / Abort edge instance
    rtrReset     : R_TRIG;                        // 复位沿检测实例 / Reset edge instance
    tonPrep      : TON;                           // 预焊段计时实例 / Pre-weld stage timer
    tonFull      : TON;                           // 满焊段计时实例 / Full-weld stage timer
    tonCrater    : TON;                           // 收弧段计时实例 / Crater stage timer
    bCfgOk       : BOOL;                          // 配方组态合法标志 / Recipe configuration valid
    bTimeOk      : BOOL;                          // 段驻留时间合法标志 / Stage dwell time valid
    nSegPrev     : INT;                           // 上一拍段号，用于冻结判据 / Previous stage for freeze criterion
    nI           : INT;                           // 配方校验循环下标 / Recipe check loop index
    uFault       : UDINT;                         // 锁存故障码，0 = 无 / Latched fault code
    uInfo        : UDINT;                         // 信息级码，永不置 bError / Info code, never raises bError
END_VAR
VAR CONSTANT
    DL_LWPS_SEGMAX : INT := 3;                    // 段总数 [段]，与数组上界一致 / Stage count matching array bound
    DL_LWPS_CNTMAX : INT := 32000;                // 冻结拍计数上限 [拍]，防 INT 溢出 / Freeze counter ceiling
END_VAR

(* === 段 0 · 实例刷新（无条件周期调用，禁入 CASE 分支）=== *)
rtrStart(CLK := bStart);                          // 每拍刷新启动沿 / Refresh start edge every scan
rtrAbort(CLK := bAbort);                          // 每拍刷新中止沿 / Refresh abort edge every scan
rtrReset(CLK := bReset);                          // 每拍刷新复位沿 / Refresh reset edge every scan
tonPrep(IN := (_eState = E_DL_LwpsPhase.ePrep), PT := atSegTime[1]);   // 预焊段计时，无条件刷新
tonFull(IN := (_eState = E_DL_LwpsPhase.eFull), PT := atSegTime[2]);   // 满焊段计时，无条件刷新
tonCrater(IN := (_eState = E_DL_LwpsPhase.eCrater), PT := atSegTime[3]); // 收弧段计时，无条件刷新

(* === 段 1 · 组态闸（每拍重算，出厂即报码，禁运行时钳位掩盖）=== *)
bCfgOk := (fRatedPowerW > fEps) AND (fDefocusMax > fEps) AND (fRatedPowerW < 1.0E7)
          AND (fRatedPowerW = fRatedPowerW) AND (fDefocusMax = fDefocusMax);   // 额定值域闸 + NaN 自反判据
bTimeOk := TRUE;                                  // 时间域先置真，逐段否决 / Assume valid then veto per stage
FOR nI := 1 TO DL_LWPS_SEGMAX DO
    bTimeOk := bTimeOk AND (atSegTime[nI] > T#0MS);                                  // 段驻留时间必须 > 0
    bCfgOk := bCfgOk AND (afSegPowerW[nI] > fEps)                                     // 功率正域闸，防 0 功率空烧
              AND (afSegPowerW[nI] <= fRatedPowerW + fEps)                            // 不超额定，防过载
              AND (afSegSpeed[nI] > fEps)                                             // 速度正域闸
              AND (ABS(afSegDefocus[nI]) <= fDefocusMax + fEps)                       // 离焦幅值域闸
              AND (afSegPowerW[nI] = afSegPowerW[nI])                                 // 功率 NaN 自反判据
              AND (afSegSpeed[nI] = afSegSpeed[nI])                                   // 速度 NaN 自反判据
              AND (afSegDefocus[nI] = afSegDefocus[nI]);                              // 离焦 NaN 自反判据
END_FOR
IF NOT bCfgOk THEN
    uFault := 16#0002_0680;                       // 故障级：配方越界，组态闸锁存
END_IF
IF NOT bTimeOk THEN
    uFault := 16#0002_0690;                       // 故障级：段驻留时间为 0，计时器无效
END_IF
uInfo := 16#0000;                                 // 信息码每拍清零，条件满足再置 / Clear info code each scan
IF nFreezeCount > 0 THEN
    uInfo := 16#0002_06A0;                        // 信息级：冻结拍已发生（不置 bError）
END_IF

(* === 段 2 · 主状态机（ENUM + CASE，含 ELSE 兜底）=== *)
CASE _eState OF
E_DL_LwpsPhase.eIdle :
    nSegNow := 0;                                 // 段号 0 = 未运行
    bSeqDone := FALSE;                            // 新一轮启动前清完成标志
    IF rtrReset.Q THEN
        uFault := 16#0000;                        // 故障产生态内提供清零点（复位路径可达）
    END_IF
    IF rtrStart.Q AND (uFault = 16#0000) THEN     // 无故障才允许启动
        _eState := E_DL_LwpsPhase.ePrep;
        nFreezeCount := 0;                        // 新序列清零冻结计数
    ELSIF uFault <> 16#0000 THEN
        _eState := E_DL_LwpsPhase.eFault;
    END_IF

E_DL_LwpsPhase.ePrep :
    nSegNow := 1;                                 // 预焊段
    bSeqDone := FALSE;
    IF tonPrep.Q THEN
        _eState := E_DL_LwpsPhase.eFull;          // 本拍行为：计时到，本拍末转满焊
    END_IF

E_DL_LwpsPhase.eFull :
    nSegNow := 2;                                 // 满焊段
    bSeqDone := FALSE;
    IF tonFull.Q THEN
        _eState := E_DL_LwpsPhase.eCrater;        // 转入收弧段
    END_IF

E_DL_LwpsPhase.eCrater :
    nSegNow := 3;                                 // 收弧段
    bSeqDone := FALSE;
    IF tonCrater.Q THEN
        _eState := E_DL_LwpsPhase.eDone;          // 收弧完成，转完成态
        bSeqDone := TRUE;                         // 置位型标志，同拍/段尾均不清零
    END_IF

E_DL_LwpsPhase.eDone :
    nSegNow := 0;                                 // 出光结束，段号归 0
    bSeqDone := TRUE;                             // 完成标志保持到下次启动
    IF rtrStart.Q OR rtrReset.Q THEN
        _eState := E_DL_LwpsPhase.eIdle;          // 再次启动或复位回空闲
    END_IF

E_DL_LwpsPhase.eFault :
    nSegNow := 0;                                 // 故障态强制段号 0（安全侧）
    IF rtrReset.Q AND bCfgOk AND bTimeOk THEN
        uFault := 16#0000;                        // 组态修正且复位沿才解锁
        _eState := E_DL_LwpsPhase.eIdle;
    END_IF

ELSE
    _eState := E_DL_LwpsPhase.eFault;             // 非法状态拦截，落故障态
    nSegNow := 0;                                 // 安全侧段号
    uFault := 16#0002_0690;                       // 故障级：段序号越界（枚举兜底路径）
END_CASE
IF rtrAbort.Q OR (NOT bEnable) THEN
    _eState := E_DL_LwpsPhase.eIdle;              // 中止/失能优先回空闲，安全侧最高优先
    nSegNow := 0;                                 // 段号随之为 0
    bSeqDone := FALSE;                            // 完成标志随之中止
END_IF

(* === 段 3 · 输出映射（安全三行同向：驱动方向 → 记账符号 → 到位判据）=== *)
IF nSegNow <> nSegPrev THEN
    nFreezeCount := nFreezeCount + 1;             // 段切换当拍：冻结输出，沿用上一拍指令
    IF nFreezeCount > DL_LWPS_CNTMAX THEN
        nFreezeCount := DL_LWPS_CNTMAX;           // 冻结计数饱和，防 INT 溢出
    END_IF
ELSE
    IF (nSegNow >= 1) AND (nSegNow <= DL_LWPS_SEGMAX) THEN
        fPowerCmdW  := afSegPowerW[nSegNow];      // 段号已钳域，数组访问安全
        fSpeedCmd   := afSegSpeed[nSegNow];       // 速度随段切换
        fDefocusCmd := afSegDefocus[nSegNow];     // 离焦随段切换
    ELSE
        fPowerCmdW  := 0.0;                       // 非运行态功率指令 0（驱动方向安全）
        fSpeedCmd   := 0.0;                       // 速度指令 0
        fDefocusCmd := 0.0;                       // 离焦指令 0
    END_IF
END_IF
bWeldActive := (nSegNow >= 1) AND (nSegNow <= DL_LWPS_SEGMAX) AND (fPowerCmdW > fEps);  // 出光判据与功率同向
nSegPrev := nSegNow;                              // 段号记账：本拍末更新，供下一拍冻结判据
bError := (uFault <> 16#0000);                    // 故障标志仅由故障级码置位（R45 配对）
IF bError THEN
    uErrorId := uFault;                           // 故障级码优先上报
ELSE
    uErrorId := uInfo;                            // 无故障时上报信息级码
END_IF
eStateOut := _eState;                             // 输出枚举段尾单点映射（N2 规则）
END_FUNCTION_BLOCK

(* ---- FB_DL_LehrZoneTempSeq.st ---- *)
(*
  Name: FB_DL_LehrZoneTempSeq
  Category: DL_Process
  Version: 1.0.0
  Round: R90 / 2026-11-25
  开源溯源：clean-room 自研（族 浮法玻璃锡槽退火，ST 开源生态实测 0 命中，无外部代码引入）
  功能：1) 退火窑分区温度时序给定：斜坡相按设定升温/降温速率把温度给定从当前保持值斜坡推到
           设定值 fSetC，到达后进保温相；保温相保持 fHoldS 后置完成位并停在保持相。
           斜坡步进按「速率 × 扫描周期」逐拍累加：ΔT = 速率[°C/min] × (周期[s]/60)，
           因此必须把扫描周期作为入参并对它做零闸（R21），不许假设固定扫描周期。
        2) 温度给定的起点是本件自身的保持值 _fOutC：完成相保持在 fSetC，再次启动即从 fSetC
           重新斜坡到新设定值，语义自洽；上电首次运行为 0 °C 起始（保持变量默认值）。
        3) 超温保护：斜坡与保温两相内，只要温度给定超过 fOverLimitC 立即进故障相并锁存，
           同时把温度给定回退到超温前的安全值（不超过上限），输出侧不再继续推高。
  边界条件：1) 非有限值闸：设定值、速率、超温上限、扫描周期四路实值入参统一过
           NOT(x > -DL_BIG AND x < DL_BIG)，同时拦 NaN 与 Inf；命中即判组态非法并进故障相，
           绝不把 NaN 累加进温度给定（一旦累加，保持值会被永久污染，R19）。
        2) 组态零闸：ABS(fCycleS) > DL_EPS 才允许积分（周期为零则斜坡不推进，且 ΔT 会除零）；
           fRateCmin 必须 > DL_EPS（速率为 0 时永远到不了设定值，属组态错误）；
           fOverLimitC 必须 > fSetC（超温上限低于设定值时保护恒动作，属组态错误）。
        3) 时间零闸：fHoldS <= T#0S 时保温相定时器立即置 Q（等价于跳过保温），
           这是合法组态（调试用），语义在此声明。
        4) 相超时说明：eLztRamp 的超时由「斜坡是否推进」间接体现（速率与周期已闸），
           另设 tonRampOv 兜底防组态导致的永久不达；eLztHold 由 tonHold 定时，无额外超时；
           eLztDone 为稳态持留相（等 xStart 撤令），不设超时。
        5) 状态机兜底：CASE 全态覆盖 + ELSE 强制回故障相；故障解除路径为
           (NOT xStart) AND 组态恢复，可达。
        6) FB 主体不使用 RETURN，统一单出口（跨平台可移植性）。
  量纲自证：ΔT = (°C/min) × (s / 60 (s/min)) = °C，步进与温度同量纲；
           fOutC = °C + °C = °C；与 fOverLimitC 同为 °C 后方可比较；
           tonXxx 的 PT 均为 [TIME]；本件无跨量纲相加。
  码表 Error codes（本件格 0090_06xx，故障级一律 3 行内置 _uFault/_bFault/_eState）:
    16#0090_0601 故障级：组态非法（周期为零/速率非正/超温上限不高于设定值/非有限）
    16#0090_0602 故障级：超温保护动作（温度给定超过上限）
    16#0090_0603 故障级：斜坡相超时兜底（长时间未到达设定值）
    16#0090_0604 故障级：状态机落 ELSE 兜底（非法相位 ID）
    16#0090_0605 信息级：斜坡已到达设定值，转入保温

  修订历史 Revision :
    2026-11-25  v1.0.0  R90 首版
*)

TYPE E_DL_LztState :
(
    eLztIdle := 0,    // 待机：等启动上升沿 / Idle, awaiting start edge
    eLztRamp := 10,   // 斜坡：按速率推向设定值 / Ramping toward setpoint
    eLztHold := 20,   // 保温：等保温时长 / Holding for the hold duration
    eLztDone := 30,   // 完成：给定保持，等撤令 / Done, setpoint held until release
    eLztFault:= 90    // 故障：锁存待解除 / Fault, latched awaiting release
);
END_TYPE

FUNCTION_BLOCK FB_DL_LehrZoneTempSeq
VAR_INPUT
    xStart      : BOOL;    // 时序启动指令（上升沿有效）[bool] / Sequence start, edge triggered [bool]
    fSetC       : REAL;    // 目标设定温度 [°C] / Target setpoint temperature [°C]
    fRateCmin   : REAL;    // 升温/降温速率 [°C/min] / Ramp rate [°C/min]
    fHoldS      : TIME;    // 保温时长 [TIME] / Hold duration [TIME]
    fOverLimitC : REAL;    // 超温保护上限 [°C] / Over-temperature protection limit [°C]
    fCycleS     : REAL;    // 扫描周期 [s] / Scan cycle time [s]
END_VAR
VAR_OUTPUT
    fOutC       : REAL;    // 温度给定输出 [°C] / Temperature setpoint output [°C]
    xDone       : BOOL;    // 时序完成保持位 [bool] / Sequence complete held flag [bool]
    xBusy       : BOOL;    // 时序进行中 [bool] / Sequence busy flag [bool]
    eState      : E_DL_LztState;   // 状态出口，段尾单点映射 / State outlet, single-point mapped
    nErrId      : UDINT;   // 事件码，0 = 无事件 / Event code, 0 = none
END_VAR
VAR
    tonHold     : TON;     // 保温时长定时器 [TIME] / Hold duration timer
    tonRampOv   : TON;     // 斜坡相超时兜底定时器 [TIME] / Ramp overrun watchdog timer
    rtStart     : R_TRIG;  // 启动上升沿检测 [bool] / Start rising edge detector
    _eState     : E_DL_LztState := E_DL_LztState.eLztIdle;   // 内部相位（CASE 唯一写入目标）
    _eStatePrev : E_DL_LztState := E_DL_LztState.eLztIdle;   // 上一拍相位快照（周期末更新）
    _fOutC      : REAL;    // 温度给定保持值 [°C] / Retained setpoint value [°C]
    _fStepC     : REAL;    // 单拍温度步进量 [°C] / Temperature step per cycle [°C]
    _bCfgBad    : BOOL;    // 组态非法聚合 [bool] / Configuration invalid aggregate [bool]
    _bAtSet     : BOOL;    // 已达设定值（带死区）[bool] / Reached setpoint within deadband [bool]
    _bOverTemp  : BOOL;    // 超温条件成立 [bool] / Over-temperature condition [bool]
    _bBusy      : BOOL;    // 激活相（斜坡/保温）[bool] / Active phase flag [bool]
    _bFault     : BOOL;    // 故障锁存位 [bool] / Latched fault flag [bool]
    _uInfo      : UDINT;   // 信息码，每拍重算 / Info code, recomputed every cycle
    _uFault     : UDINT;   // 故障码锁存 / Latched fault code
END_VAR
VAR CONSTANT
    DL_EPS      : REAL := 1.0E-9;    // 组态零闸阈值 [-] / Configuration zero gate threshold [-]
    DL_BIG      : REAL := 1.0E12;    // 非有限值闸量级上限 [-] / Finiteness gate magnitude [-]
    DL_S_PER_MIN: REAL := 60.0;      // min → s 换算因子 [s/min] / Minute to second factor [s/min]
    DL_DEADBAND : REAL := 0.05;      // 到达设定值的死区 [°C] / Setpoint arrival deadband [°C]
    DL_RAMP_MAX : TIME := T#4H;      // 斜坡相超时兜底上限 [TIME] / Ramp overrun ceiling [TIME]
END_VAR

(* —— 段 0：单拍量预清零（锁存量 _uFault/_bFault/_fOutC/_eStatePrev 不入清单，R187①） —— *)
_uInfo := 16#0000_0000;                     // 信息码每拍重算 / Info code recomputed
nErrId := 16#0000_0000;                     // 事件码缺省无事件 / Event code defaults to none

(* —— 段 1：非有限值闸（R19：NaN 一旦累加进保持值会永久污染，必须前置拦截） —— *)
_bCfgBad := NOT (fSetC > -DL_BIG AND fSetC < DL_BIG)
            OR NOT (fRateCmin > -DL_BIG AND fRateCmin < DL_BIG)
            OR NOT (fOverLimitC > -DL_BIG AND fOverLimitC < DL_BIG)
            OR NOT (fCycleS > -DL_BIG AND fCycleS < DL_BIG);

(* —— 段 2：组态零闸（R4 / R21：周期与速率两个零闸，另加超温上限的逻辑闸） —— *)
_bCfgBad := _bCfgBad
            OR (ABS(fCycleS) <= DL_EPS)               // 周期为零：积分不推进且步进发散
            OR (fRateCmin <= DL_EPS)                  // 速率为零：永远到不了设定值
            OR (fOverLimitC <= fSetC)                 // 超温上限不高于设定值：保护恒动作
            OR (fRateCmin > DL_BIG);                  // 速率荒谬：拒绝进入运算

(* —— 段 3：步进量与判据量（每拍重算） —— *)
IF _bCfgBad THEN
    _fStepC := 0.0;                               // 组态坏：步进量置 0，保持值不动
ELSE
    _fStepC := fRateCmin * (fCycleS / DL_S_PER_MIN);   // 速率 × 周期 = 单拍步进 [°C]
END_IF
_bAtSet := (NOT _bCfgBad) AND (ABS(fSetC - _fOutC) <= DL_DEADBAND);   // 已达设定值
_bOverTemp := (NOT _bCfgBad) AND (_fOutC > fOverLimitC);              // 超温条件

(* —— 段 4：激活量与定时器无条件周期刷新（R7：调用语句不得置于 IF/CASE 内） —— *)
_bBusy := (_eState = E_DL_LztState.eLztRamp) OR (_eState = E_DL_LztState.eLztHold);
rtStart(CLK := xStart);                                                  // 启动上升沿，每拍必调
tonHold(IN := (_eState = E_DL_LztState.eLztHold), PT := fHoldS);         // 保温时长
tonRampOv(IN := (_eState = E_DL_LztState.eLztRamp), PT := DL_RAMP_MAX);  // 斜坡超时兜底

(* —— 段 5：全局故障拦截（优先级最高；已锁存则不再改写码值，禁同拍抹除） —— *)
IF _bCfgBad AND (NOT _bFault) THEN
    _uFault := 16#0090_0601;                // 故障级：组态非法
    _bFault := TRUE;                        // 锁存（3 行内置，R45 配对）
    _eState := E_DL_LztState.eLztFault;
END_IF
IF _bOverTemp AND _bBusy AND (NOT _bFault) THEN
    _uFault := 16#0090_0602;                // 故障级：超温保护动作
    _bFault := TRUE;                        // 锁存
    _eState := E_DL_LztState.eLztFault;
END_IF
IF tonRampOv.Q AND (_eState = E_DL_LztState.eLztRamp) AND (NOT _bFault) THEN
    _uFault := 16#0090_0603;                // 故障级：斜坡相超时兜底
    _bFault := TRUE;                        // 锁存
    _eState := E_DL_LztState.eLztFault;
END_IF

(* —— 段 6：相位机与斜坡积分（只做迁移与保持值更新；出口在段 8 单点映射） —— *)
CASE _eState OF

E_DL_LztState.eLztIdle:
    IF NOT xStart THEN
        ;                                   // 等启动，保持值不变 / Waiting, retained value held
    ELSIF rtStart.Q THEN
        _eState := E_DL_LztState.eLztRamp;  // 进斜坡相
    END_IF

E_DL_LztState.eLztRamp:
    IF NOT xStart THEN
        _eState := E_DL_LztState.eLztIdle;  // 撤令：回待机（保持值保留）
    ELSIF _bAtSet THEN
        _uInfo := 16#0090_0605;             // 信息级：已到达设定值
        _eState := E_DL_LztState.eLztHold;  // 进保温相
    ELSE
        IF _fOutC < fSetC THEN
            _fOutC := MIN(fSetC, _fOutC + _fStepC);   // 升温：向上逼近，不越过设定值
        ELSE
            _fOutC := MAX(fSetC, _fOutC - _fStepC);   // 降温：向下逼近，不越过设定值
        END_IF
    END_IF

E_DL_LztState.eLztHold:
    IF NOT xStart THEN
        _eState := E_DL_LztState.eLztIdle;  // 撤令：回待机
    ELSIF tonHold.Q THEN
        _eState := E_DL_LztState.eLztDone;  // 保温结束：进完成相
    END_IF

E_DL_LztState.eLztDone:
    IF _bOverTemp THEN
        ;                                   // 超温由段 5 全局拦截，此处不重复赋值
    ELSIF NOT xStart THEN
        _eState := E_DL_LztState.eLztIdle;  // 撤令：回待机
    END_IF

E_DL_LztState.eLztFault:
    IF (NOT xStart) AND (NOT _bCfgBad) THEN
        _bFault := FALSE;                   // 解除路径：撤令 + 组态恢复（可达）
        _uFault := 16#0000_0000;            // 清锁存码
        _eState := E_DL_LztState.eLztIdle;  // 回待机
    END_IF

ELSE
    _uFault := 16#0090_0604;                // 故障级：非法相位 ID 兜底
    _bFault := TRUE;                        // 锁存
    _eState := E_DL_LztState.eLztFault;     // 强制回故障相

END_CASE

(* —— 段 7：后置段（R23：保持值安全回退与快照统一放在迁移判断之后） —— *)
IF _fOutC > fOverLimitC THEN
    _fOutC := fOverLimitC;                  // 超温回退：保持值不得高于上限（安全侧）
END_IF
_eStatePrev := _eState;                     // 快照统一在周期末尾更新（R23）

(* —— 段 8：出口单点映射（名实同源；由状态与保持值导出，不在多分支各写一遍） —— *)
fOutC := _fOutC;                                              // 温度给定出口 [°C]
xBusy := _bBusy AND (NOT _bFault);                            // 进行中出口
xDone := (_eState = E_DL_LztState.eLztDone) AND (NOT _bFault); // 完成位出口
eState := _eState;                                            // 状态出口单点映射
IF _bFault THEN
    nErrId := _uFault;                      // 故障锁存码回放（不在故障相按当下输入重推断）
ELSE
    nErrId := _uInfo;                       // 信息码
END_IF

END_FUNCTION_BLOCK
